(* IEC 61131-3 sources: volt/packages/volt-lsp-iec/test-corpus/awa-palletizer/Device/Plc Logic/Application/Library Manager/L_UMTP_Mathematics, 222 files *)

(* ---- L_UMTP_COMPLEX.dut ---- *)
TYPE L_UMTP_COMPLEX :
STRUCT
	LRRE : LREAL;
	LRIM : LREAL;
END_STRUCT
END_TYPE

(* ---- L_UMTP_INTERPOLATIONDATA.dut ---- *)
TYPE L_UMTP_INTERPOLATIONDATA :
STRUCT
	PARRX : POINTER TO LREAL;
	XISEQUIDISTANT : BOOL;
	UDISTRIDEX : UDINT;
	PARRY : POINTER TO LREAL;
	YISEQUIDISTANT : BOOL;
	UDISTRIDEY : UDINT;
	UICOUNT : UDINT;
	OPTIONS : UDINT;
END_STRUCT
END_TYPE

(* ---- L_UMTP_INTERPOLATIONTYPE.dut ---- *)
TYPE L_UMTP_INTERPOLATIONTYPE :
(
	UNDEFINED := 0,
	LINEAR := 1,
	CUBICSPLINENATURAL := 30,
	CUBICSPLINEHERMITE := 31,
	CUBICSPLINEHERMITEEXTERN := 32,
	NEWTON := 5
);
END_TYPE

(* ---- L_UMTP_MATRIX3X3.dut ---- *)
TYPE L_UMTP_MATRIX3X3 :
STRUCT
	M11 : LREAL;
	M12 : LREAL;
	M13 : LREAL;
	M21 : LREAL;
	M22 : LREAL;
	M23 : LREAL;
	M31 : LREAL;
	M32 : LREAL;
	M33 : LREAL;
END_STRUCT
END_TYPE

(* ---- L_UMTP_QUATERNION.dut ---- *)
TYPE L_UMTP_QUATERNION :
STRUCT
	LRRE : LREAL;
	LRIM1 : LREAL;
	LRIM2 : LREAL;
	LRIM3 : LREAL;
END_STRUCT
END_TYPE

(* ---- L_UMTP_REVERSEPOLISHNOTATIONTOKEN.dut ---- *)
TYPE L_UMTP_REVERSEPOLISHNOTATIONTOKEN :
(
	NONE := 0,
	PARENTHESIS := 1,
	FLOAT := 2,
	BOOLEAN := 3,
	NEGOTIATE := 4,
	PLUS := 10,
	MINUS := 11,
	MULTIPLIKATION := 12,
	DIVISION := 13,
	POW := 14,
	MODULO := 15,
	SINE := 20,
	COSINE := 21,
	TANGENS := 22,
	ASINE := 23,
	ACOSINE := 24,
	ATANGENS := 25,
	EXPONENTIAL := 40,
	LOGN := 41,
	LOG10 := 42,
	SQUAREROOT := 43,
	ABSOLUTE := 44,
	SIGNUM := 45,
	CEIL := 50,
	FLOOR := 51,
	TRUNCATE := 52,
	ROUND := 53,
	EQUAL := 100,
	NOTEQUAL := 101,
	GREATEREQUAL := 102,
	GREATERTHEN := 103,
	LESSEQUAL := 104,
	LESSTHEN := 105,
	LOGICAND := 110,
	LOGICXOR := 111,
	LOGICOR := 112,
	LOGICNOT := 113
);
END_TYPE

(* ---- L_UMTP_ROBOTACC.dut ---- *)
TYPE L_UMTP_ROBOTACC :
STRUCT
	ACC : L_UMTP_Vector3D;
	PITCH : L_UMTP_Vector3D;
END_STRUCT
END_TYPE

(* ---- L_UMTP_ROBOTFRAME.dut ---- *)
TYPE L_UMTP_ROBOTFRAME :
STRUCT
	POS : L_UMTP_RobotPos;
	VEL : L_UMTP_RobotVel;
	ACC : L_UMTP_RobotAcc;
END_STRUCT
END_TYPE

(* ---- L_UMTP_ROBOTPOS.dut ---- *)
TYPE L_UMTP_ROBOTPOS :
STRUCT
	POS : L_UMTP_Vector3D;
	ROT : L_UMTP_RotMat;
END_STRUCT
END_TYPE

(* ---- L_UMTP_ROBOTVEL.dut ---- *)
TYPE L_UMTP_ROBOTVEL :
STRUCT
	VEL : L_UMTP_Vector3D;
	TWIST : L_UMTP_Vector3D;
END_STRUCT
END_TYPE

(* ---- L_UMTP_ROTATIONCONVENTION.dut ---- *)
TYPE L_UMTP_ROTATIONCONVENTION :
(
	XYZ_ROTATED := 0,
	ZYX_ROTATED := 1,
	XZY_ROTATED := 2,
	YZX_ROTATED := 3,
	YXZ_ROTATED := 4,
	ZXY_ROTATED := 5,
	XYZ_FIXED := 100,
	ZYX_FIXED := 101,
	XZY_FIXED := 102,
	YZX_FIXED := 103,
	YXZ_FIXED := 104,
	ZXY_FIXED := 105
);
END_TYPE

(* ---- L_UMTP_ROTMAT.dut ---- *)
TYPE L_UMTP_ROTMAT :
STRUCT
	PARAM : L_UMTP_RotParam;
END_STRUCT
END_TYPE

(* ---- L_UMTP_ROTPARAM.dut ---- *)
TYPE L_UMTP_ROTPARAM :
STRUCT
	SINA : LREAL;
	COSA : LREAL;
	SINB : LREAL;
	COSB : LREAL;
	SINC : LREAL;
	COSC : LREAL;
	EROTCON : L_UMTP_RotationConvention;
	XGIMBALLOCK : BOOL;
END_STRUCT
END_TYPE

(* ---- L_UMTP_TRIGONOMETRICUNIT.dut ---- *)
TYPE L_UMTP_TRIGONOMETRICUNIT :
(
	RADIANT := 0,
	DEGREE := 1
);
END_TYPE

(* ---- L_UMTP_VALIDLREAL.dut ---- *)
TYPE L_UMTP_VALIDLREAL :
STRUCT
	XVALID : BOOL;
	LRVALUE : LREAL;
END_STRUCT
END_TYPE

(* ---- L_UMTP_VECTOR3D.dut ---- *)
TYPE L_UMTP_VECTOR3D :
STRUCT
	X : LREAL;
	Y : LREAL;
	Z : LREAL;
END_STRUCT
END_TYPE

(* ---- L_UMTP_CONSTANTS.gvl ---- *)
VAR_GLOBAL
	GC_CTRLPTMAXNR : INT := 200;
	GC_IMAXNUMOFGIVENPTS : INT := 199;
	GC_UDIMAXCUBSPLINEPTS : UDINT := 11;
	G_MAXPATHDIM : DINT := 8;
	GCDWSIZEOFLREAL : DWORD := USINT_TO_DWORD(SIZEOF(LREAL));
END_VAR

(* ---- L_UMTP_DEFINES.gvl ---- *)
VAR_GLOBAL
	G_XOPTIMIZEDFRAMECALC : BOOL := TRUE;
END_VAR

(* ---- L_UMTP_MATH.gvl ---- *)
VAR_GLOBAL
	RAD2DEG : LREAL := (180.0 / Math.PI);
	DEG2RAD : LREAL := (Math.PI / 180.0);
	GRAVITY_MM : LREAL := (9.81 * 1000.0);
	EPS_REAL : LREAL := 1E-06;
	GC_LREPSILON : LREAL := 1E-09;
	EPS_LREAL : LREAL := 1E-12;
	MM2M : LREAL := 0.001;
	M2MM : LREAL := 1000;
	GCGIMBALLOCKTOL : LREAL := 5E-05;
	GCLRINVPI : LREAL := (1 / MATH.PI);
	GCLR2PI : LREAL := (2 * MATH.PI);
	GCLRINV2PI : LREAL := (1 / (2 * MATH.PI));
	GCLRPIHALF : LREAL := (MATH.PI / 2);
	GCLRINVPIHALF : LREAL := (1 / (MATH.PI / 2));
	MAXDOUBLE : LREAL := 1.79769E+308;
	MINDOUBLE : LREAL := -1.79769E+308;
	GC_POSITIVE_LIMIT_16BIT_LREAL : LREAL := 65535.0;
	GC_POSITIVE_LIMIT_15BIT_LREAL : LREAL := 32767.0;
	GC_NEGATIVE_LIMIT_15BIT_LREAL : LREAL := -32768.0;
	GC_POSITIVE_LIMIT_32BIT : LREAL := 2147483647;
	GC_NEGATIVE_LIMIT_32BIT : LREAL := -2147483647;
	GC_POSITIVE_LIMIT_32BIT_LREAL : LREAL := 4294967296.0;
	GC_POSITIVE_LIMIT_31BIT_LREAL : LREAL := 2147483647.0;
	GC_NEGATIVE_LIMIT_31BIT_LREAL : LREAL := -2147483648.0;
	GC_POSITIVE_LIMIT_63BIT_LREAL : LREAL := 9.2233720368547758E+18;
	GC_NEGATIVE_LIMIT_63BIT_LREAL : LREAL := -9.2233720368547758E+18;
	GC_POSITIVE_LIMIT_63BIT : LINT := 9223372036854775807;
	GC_NEGATIVE_LIMIT_63BIT : LINT := -9223372036854775808;
	LRCOS_0 : LREAL := 1.0;
	LRCOS_15 : LREAL := 0.965925826289068;
	LRCOS_30 : LREAL := 0.866025403784439;
	LRCOS_45 : LREAL := 0.707106781186547;
	LRCOS_60 : LREAL := 0.5;
	LRCOS_75 : LREAL := 0.258819045102521;
	LRCOS_90 : LREAL := 0.0;
	LRCOS_105 : LREAL := -0.258819045102521;
	LRCOS_120 : LREAL := -0.5;
	LRCOS_135 : LREAL := -0.707106781186548;
	LRCOS_150 : LREAL := -0.866025403784439;
	LRCOS_165 : LREAL := -0.965925826289068;
	LRCOS_180 : LREAL := -1.0;
	LRCOS_195 : LREAL := -0.965925826289068;
	LRCOS_210 : LREAL := -0.866025403784439;
	LRCOS_225 : LREAL := -0.707106781186547;
	LRCOS_240 : LREAL := -0.5;
	LRCOS_255 : LREAL := -0.258819045102521;
	LRCOS_270 : LREAL := 0.0;
	LRCOS_285 : LREAL := 0.258819045102521;
	LRCOS_300 : LREAL := 0.5;
	LRCOS_315 : LREAL := 0.707106781186548;
	LRCOS_330 : LREAL := 0.866025403784439;
	LRCOS_345 : LREAL := 0.965925826289068;
	LRCOS_360 : LREAL := 1.0;
	LRSIN_0 : LREAL := 0.0;
	LRSIN_15 : LREAL := 0.258819045102521;
	LRSIN_30 : LREAL := 0.5;
	LRSIN_45 : LREAL := 0.707106781186548;
	LRSIN_60 : LREAL := 0.866025403784439;
	LRSIN_75 : LREAL := 0.965925826289068;
	LRSIN_90 : LREAL := 1.0;
	LRSIN_105 : LREAL := 0.965925826289068;
	LRSIN_120 : LREAL := 0.866025403784439;
	LRSIN_135 : LREAL := 0.707106781186547;
	LRSIN_150 : LREAL := 0.5;
	LRSIN_165 : LREAL := 0.258819045102521;
	LRSIN_180 : LREAL := 0.0;
	LRSIN_195 : LREAL := -0.258819045102521;
	LRSIN_210 : LREAL := -0.5;
	LRSIN_225 : LREAL := -0.707106781186548;
	LRSIN_240 : LREAL := -0.866025403784439;
	LRSIN_255 : LREAL := -0.965925826289068;
	LRSIN_270 : LREAL := -1.0;
	LRSIN_285 : LREAL := -0.965925826289068;
	LRSIN_300 : LREAL := -0.866025403784439;
	LRSIN_315 : LREAL := -0.707106781186547;
	LRSIN_330 : LREAL := -0.5;
	LRSIN_345 : LREAL := -0.258819045102521;
	LRSIN_360 : LREAL := 0.0;
	L_UMTP_VALUEIGNORE : LREAL := 1E+300;
	L_UMTP_VALUEINITIAL : LREAL := 1E+301;
	L_UMTP_VALUEINVALID : LREAL := 1E+302;
	L_UMTP_VALUEINF : LREAL := 1.7976931348623157E+308;
END_VAR

(* ---- L_UMTP_FUNC_1D21D.itf ---- *)
INTERFACE L_UMTP_FUNC_1D21D
END_INTERFACE

METHOD CALL_1D21D : LREAL
VAR_INPUT
	X : LREAL;
	CONTEXT : DINT;
END_VAR
END_METHOD

(* ---- L_UMTP_FUNC_ND21D.itf ---- *)
INTERFACE L_UMTP_FUNC_ND21D
END_INTERFACE

METHOD CALL_ND21D : LREAL
VAR_INPUT
	PLRX : POINTER TO LREAL;
	UDIDIM : UDINT;
	CONTEXT : DINT;
END_VAR
END_METHOD

(* ---- L_UMTP_FUNC_ND2MD.itf ---- *)
INTERFACE L_UMTP_FUNC_ND2MD
END_INTERFACE

METHOD CALL_ND2MD
VAR_INPUT
	PLRX : POINTER TO LREAL;
	UDIXDIM : UDINT;
	PLRY : POINTER TO LREAL;
	UDIYDIM : UDINT;
	CONTEXT : DINT;
END_VAR
END_METHOD

(* ---- L_UMTP_IFFTDATA.itf ---- *)
INTERFACE L_UMTP_IFFTDATA
END_INTERFACE

METHOD RECORDDATA : UDINT
VAR_INPUT
	PLCDATA : POINTER TO L_umtp_complex;
	UDISIZEOFDATA : UDINT;
END_VAR
END_METHOD

METHOD STARTRECORDING : BOOL
END_METHOD

METHOD STOPRECORDING : BOOL
END_METHOD

(* ---- L_UMTP_IINTERPOLATION.itf ---- *)
INTERFACE L_UMTP_IINTERPOLATION
END_INTERFACE

METHOD GETVALUE : BOOL
VAR_INPUT
	X : LREAL;
END_VAR
VAR_OUTPUT
	Y : LREAL;
END_VAR
END_METHOD

(* ---- L_UMTP_IMETRIC.itf ---- *)
INTERFACE L_UMTP_IMETRIC
END_INTERFACE

METHOD DISTANCE : LREAL
VAR_INPUT
	ITFOB1 : __SYSTEM.IQueryInterface;
	ITFOB2 : __SYSTEM.IQueryInterface;
END_VAR
END_METHOD

(* ---- L_UMTP_IODE.itf ---- *)
INTERFACE L_UMTP_IODE
END_INTERFACE

METHOD FIRSTDERIV
VAR_INPUT
	PLRY : POINTER TO LREAL;
	PLRDY : POINTER TO LREAL;
	UDIDIM : UDINT;
	LRT : LREAL;
END_VAR
END_METHOD

(* ---- L_UMTP_IPATH.itf ---- *)
INTERFACE L_UMTP_IPATH
END_INTERFACE

METHOD GETPATHVALUE : BOOL
VAR_INPUT
	PLRX : POINTER TO LREAL;
	PLRD1 : POINTER TO LREAL;
	PLRD2 : POINTER TO LREAL;
	UDIDIM : UDINT;
	LRU : LREAL;
END_VAR
END_METHOD

(* ---- L_UMTP_ISORTDATA.itf ---- *)
INTERFACE L_UMTP_ISORTDATA
END_INTERFACE

METHOD EXCHANGE : BOOL
VAR_INPUT
	IDX1 : DINT;
	IDX2 : DINT;
END_VAR
END_METHOD

METHOD GETVALUE : LREAL
VAR_INPUT
	IDX : DINT;
END_VAR
END_METHOD

(* ---- CALCCARTLENGTH.pou ---- *)
FUNCTION CALCCARTLENGTH : LREAL
VAR_INPUT
	PVEC : POINTER TO LREAL;
	NUMELEMENTS : __XWORD;
END_VAR
END_FUNCTION

(* ---- CAPITAL_CASE.pou ---- *)
FUNCTION CAPITAL_CASE : STRING(255)
VAR_INPUT
	STR : STRING(255);
END_VAR
END_FUNCTION

(* ---- DELETE_FROM_STR.pou ---- *)
FUNCTION DELETE_FROM_STR : STRING(255)
VAR_INPUT
	STR1 : STRING(255);
	STR2 : STRING(255);
END_VAR
END_FUNCTION

(* ---- GETBOOLEANPROPERTY.pou ---- *)
FUNCTION GETBOOLEANPROPERTY : BOOL
VAR_INPUT
	STKEY : WSTRING;
END_VAR
END_FUNCTION

(* ---- GETCOMPANY.pou ---- *)
FUNCTION GETCOMPANY : WSTRING
END_FUNCTION

(* ---- GETNUMBERPROPERTY.pou ---- *)
FUNCTION GETNUMBERPROPERTY : DINT
VAR_INPUT
	STKEY : WSTRING;
END_VAR
END_FUNCTION

(* ---- GETTEXTPROPERTY.pou ---- *)
FUNCTION GETTEXTPROPERTY : WSTRING
VAR_INPUT
	STKEY : WSTRING;
END_VAR
END_FUNCTION

(* ---- GETTEXTPROPERTY2.pou ---- *)
FUNCTION GETTEXTPROPERTY2 : POINTER TO WSTRING
VAR_INPUT
	STKEY : WSTRING;
END_VAR
END_FUNCTION

(* ---- GETTITLE.pou ---- *)
FUNCTION GETTITLE : WSTRING
END_FUNCTION

(* ---- GETVERSION.pou ---- *)
FUNCTION GETVERSION : VERSION
END_FUNCTION

(* ---- GETVERSIONPROPERTY.pou ---- *)
FUNCTION GETVERSIONPROPERTY : VERSION
VAR_INPUT
	STKEY : WSTRING;
END_VAR
END_FUNCTION

(* ---- L_UMTP_2DINTERPOLATIONLINEAR.pou ---- *)
FUNCTION L_UMTP_2DINTERPOLATIONLINEAR : BOOL
VAR_INPUT
	ALRX : POINTER TO LREAL;
	ALRY : POINTER TO LREAL;
	ALRZ : POINTER TO LREAL;
	LRX : LREAL;
	LRY : LREAL;
END_VAR
VAR_OUTPUT
	XERROR : BOOL;
	EERRORID : L_IE1P_Error;
	LRZ : LREAL;
END_VAR
END_FUNCTION

(* ---- L_UMTP_ABC2ROT.pou ---- *)
FUNCTION L_UMTP_ABC2ROT
VAR_INPUT
	ROTMAT : REFERENCE TO L_UMTP_RotMat;
END_VAR
END_FUNCTION

(* ---- L_UMTP_ANTISYMTIMESMATRIX3D.pou ---- *)
FUNCTION L_UMTP_ANTISYMTIMESMATRIX3D
VAR_INPUT
	M : REFERENCE TO L_UMTP_Matrix3x3;
	TWIST : REFERENCE TO L_UMTP_Vector3D;
	RESULT : REFERENCE TO L_UMTP_Matrix3x3;
END_VAR
END_FUNCTION

(* ---- L_UMTP_APPENDPITCH.pou ---- *)
FUNCTION L_UMTP_APPENDPITCH : BOOL
VAR_INPUT
	DPHIA : LREAL;
	DPHIB : LREAL;
	DPHIC : LREAL;
	DDPHIA : LREAL;
	DDPHIB : LREAL;
	DDPHIC : LREAL;
	FRAME : REFERENCE TO L_UMTP_RobotFrame;
END_VAR
END_FUNCTION

(* ---- L_UMTP_APPENDTWIST.pou ---- *)
FUNCTION L_UMTP_APPENDTWIST : BOOL
VAR_INPUT
	DPHIA : LREAL;
	DPHIB : LREAL;
	DPHIC : LREAL;
	FRAME : REFERENCE TO L_UMTP_RobotFrame;
END_VAR
END_FUNCTION

(* ---- L_UMTP_APPROXSIGN.pou ---- *)
FUNCTION L_UMTP_APPROXSIGN : LREAL
VAR_INPUT
	LRX : LREAL;
	LRFAC : LREAL;
END_VAR
END_FUNCTION

(* ---- L_UMTP_ATAN2.pou ---- *)
FUNCTION L_UMTP_ATAN2 : LREAL
VAR_INPUT
	LRSINUS : LREAL;
	LRCOSINUS : LREAL;
END_VAR
END_FUNCTION

(* ---- L_UMTP_BENDING.pou ---- *)
FUNCTION L_UMTP_BENDING : LREAL
VAR_INPUT
	ALRD1 : REFERENCE TO ARRAY [1..3] OF LREAL;
	ALRD2 : REFERENCE TO ARRAY [1..3] OF LREAL;
END_VAR
END_FUNCTION

(* ---- L_UMTP_BILINEARINTERPOLATION.pou ---- *)
FUNCTION L_UMTP_BILINEARINTERPOLATION : BOOL
VAR_INPUT
	LRX0 : LREAL;
	LRX1 : LREAL;
	LRY0 : LREAL;
	LRY1 : LREAL;
	LRZ00 : LREAL;
	LRZ01 : LREAL;
	LRZ10 : LREAL;
	LRZ11 : LREAL;
	LRX : LREAL;
	LRY : LREAL;
END_VAR
VAR_OUTPUT
	LRZ : LREAL;
END_VAR
END_FUNCTION

(* ---- L_UMTP_BISECTION.pou ---- *)
FUNCTION L_UMTP_BISECTION : BOOL
VAR_INPUT
	IFUNC : L_UMTP_Func_1D21D;
	CONTEXT : DINT;
	A : LREAL;
	B : LREAL;
	F_REQUESTED : LREAL;
	TOL : LREAL;
	X : REFERENCE TO LREAL;
END_VAR
END_FUNCTION

(* ---- L_UMTP_BRENTALGORITHM.pou ---- *)
FUNCTION L_UMTP_BRENTALGORITHM : BOOL
VAR_INPUT
	IFUNC : L_UMTP_Func_1D21D;
	CONTEXT : DINT;
	A : LREAL;
	B : LREAL;
	TOL : LREAL;
	X : REFERENCE TO LREAL;
END_VAR
END_FUNCTION

(* ---- L_UMTP_BUBBLESORTINT.pou ---- *)
FUNCTION L_UMTP_BUBBLESORTINT
VAR_INPUT
	PIX : POINTER TO INT;
	UDISIZE : UDINT;
	XINVERT : BOOL;
END_VAR
END_FUNCTION

(* ---- L_UMTP_BUBBLESORTITFSORTDATA.pou ---- *)
FUNCTION L_UMTP_BUBBLESORTITFSORTDATA : BOOL
VAR_INPUT
	ITFDATA : L_UMTP_ISortData;
	XINVERT : BOOL;
END_VAR
END_FUNCTION

(* ---- L_UMTP_BUBBLESORTLREAL.pou ---- *)
FUNCTION L_UMTP_BUBBLESORTLREAL
VAR_INPUT
	PLRX : POINTER TO LREAL;
	UDISIZE : UDINT;
	XINVERT : BOOL;
END_VAR
END_FUNCTION

(* ---- L_UMTP_CHECKGIMBALLOCK.pou ---- *)
FUNCTION L_UMTP_CHECKGIMBALLOCK : BOOL
VAR_INPUT
	PARAM : REFERENCE TO L_UMTP_RotParam;
END_VAR
END_FUNCTION

(* ---- L_UMTP_CHECKMONOTONIC.pou ---- *)
FUNCTION L_UMTP_CHECKMONOTONIC : BYTE
VAR_INPUT
	PLRVALUES : POINTER TO LREAL;
	NDATA : UDINT;
	NSTRIDE : UDINT;
END_VAR
END_FUNCTION

(* ---- L_UMTP_CHECKSTEPSIZE.pou ---- *)
FUNCTION L_UMTP_CHECKSTEPSIZE : BOOL
VAR_INPUT
	PLRY0 : POINTER TO LREAL;
	PLRY1 : POINTER TO LREAL;
	UDIDIM : UDINT;
	LRTOL : LREAL;
	LRH : LREAL;
END_VAR
VAR_OUTPUT
	LRHTOL : LREAL;
END_VAR
END_FUNCTION

(* ---- L_UMTP_CLEAR.pou ---- *)
FUNCTION L_UMTP_CLEAR : BOOL
VAR_INPUT
	ALRARR : POINTER TO LREAL;
END_VAR
END_FUNCTION

(* ---- L_UMTP_COMEQ.pou ---- *)
FUNCTION L_UMTP_COMEQ : BOOL
VAR_INPUT
	COMVALUE : L_UMTP_Complex;
	COMTARGET : L_UMTP_Complex;
END_VAR
END_FUNCTION

(* ---- L_UMTP_COMPLEX2MAGNITUDE.pou ---- *)
FUNCTION L_UMTP_COMPLEX2MAGNITUDE : LREAL
VAR_INPUT
	SCCOIN : L_UMTP_Complex;
END_VAR
END_FUNCTION

(* ---- L_UMTP_COMPLEXCART2POLAR.pou ---- *)
FUNCTION L_UMTP_COMPLEXCART2POLAR
VAR_INPUT
	SCCOIN : L_UMTP_Complex;
	ETRIGUNIT : L_UMTP_TrigonometricUnit;
END_VAR
VAR_OUTPUT
	LRMAGNITUDE : LREAL;
	LRANGLE : LREAL;
END_VAR
END_FUNCTION

(* ---- L_UMTP_COMPLEXDIV.pou ---- *)
FUNCTION L_UMTP_COMPLEXDIV : L_UMTP_Complex
VAR_INPUT
	SCCOIN1 : L_UMTP_complex;
	SCCOIN2 : L_UMTP_complex;
END_VAR
END_FUNCTION

(* ---- L_UMTP_COMPLEXMUL.pou ---- *)
FUNCTION L_UMTP_COMPLEXMUL : L_UMTP_Complex
VAR_INPUT
	COIN1 : L_UMTP_complex;
	COIN2 : L_UMTP_complex;
END_VAR
END_FUNCTION

(* ---- L_UMTP_COMPLEXPOLAR2CART.pou ---- *)
FUNCTION L_UMTP_COMPLEXPOLAR2CART : L_UMTP_Complex
VAR_INPUT
	LRMAGNITUDE : LREAL;
	LRANGLE : LREAL;
	ETRIGUNIT : L_UMTP_TrigonometricUnit;
END_VAR
END_FUNCTION

(* ---- L_UMTP_CONFIGURATIONABC.pou ---- *)
FUNCTION L_UMTP_CONFIGURATIONABC : INT
VAR_INPUT
	ROTMAT : REFERENCE TO L_UMTP_RotMat;
END_VAR
END_FUNCTION

(* ---- L_UMTP_CROSS.pou ---- *)
FUNCTION L_UMTP_CROSS : BOOL
VAR_INPUT
	A : REFERENCE TO ARRAY [1..3] OF LREAL;
	B : REFERENCE TO ARRAY [1..3] OF LREAL;
	RESULT : REFERENCE TO ARRAY [1..3] OF LREAL;
END_VAR
END_FUNCTION

(* ---- L_UMTP_CROSSPROD.pou ---- *)
FUNCTION L_UMTP_CROSSPROD : BOOL
VAR_IN_OUT
	ALRA : ARRAY [1..3] OF LREAL;
	ALRB : ARRAY [1..3] OF LREAL;
	ALRRESULT : ARRAY [1..3] OF LREAL;
END_VAR
END_FUNCTION

(* ---- L_UMTP_DABC2DROT.pou ---- *)
FUNCTION L_UMTP_DABC2DROT
VAR_INPUT
	PARAM : REFERENCE TO L_UMTP_RotParam;
	DPHIA : LREAL;
	DPHIB : LREAL;
	DPHIC : LREAL;
	DROT : REFERENCE TO L_UMTP_Matrix3x3;
END_VAR
END_FUNCTION

(* ---- L_UMTP_DDABC2DDROT.pou ---- *)
FUNCTION L_UMTP_DDABC2DDROT
VAR_INPUT
	PARAM : L_UMTP_RotParam;
	DPHIA : LREAL;
	DPHIB : LREAL;
	DPHIC : LREAL;
	DDPHIA : LREAL;
	DDPHIB : LREAL;
	DDPHIC : LREAL;
	DDROT : REFERENCE TO L_UMTP_Matrix3x3;
END_VAR
END_FUNCTION

(* ---- L_UMTP_DDROT2DDABC.pou ---- *)
FUNCTION L_UMTP_DDROT2DDABC
VAR_INPUT
	PARAM : REFERENCE TO L_UMTP_RotParam;
	DDROT : REFERENCE TO L_UMTP_Matrix3x3;
	DPHIA : LREAL;
	DPHIB : LREAL;
	DPHIC : LREAL;
END_VAR
VAR_OUTPUT
	DDPHIA : LREAL;
	DDPHIB : LREAL;
	DDPHIC : LREAL;
END_VAR
END_FUNCTION

(* ---- L_UMTP_DDROT2FRAME.pou ---- *)
FUNCTION L_UMTP_DDROT2FRAME : BOOL
VAR_INPUT
	FRAME : REFERENCE TO L_UMTP_RobotFrame;
	DDROT : REFERENCE TO L_UMTP_Matrix3x3;
END_VAR
END_FUNCTION

(* ---- L_UMTP_DETERMINAT3D.pou ---- *)
FUNCTION L_UMTP_DETERMINAT3D : LREAL
VAR_IN_OUT
	M : L_UMTP_Matrix3x3;
END_VAR
END_FUNCTION

(* ---- L_UMTP_DISTANCE.pou ---- *)
FUNCTION L_UMTP_DISTANCE : LREAL
VAR_INPUT
	PLRX : POINTER TO LREAL;
	PLRY : POINTER TO LREAL;
	UDIDIM : UDINT;
END_VAR
END_FUNCTION

(* ---- L_UMTP_DIV.pou ---- *)
FUNCTION L_UMTP_DIV : LREAL
VAR_INPUT
	A : LREAL;
	B : LREAL;
END_VAR
END_FUNCTION

(* ---- L_UMTP_DORMANDPRINCE45STEP.pou ---- *)
FUNCTION L_UMTP_DORMANDPRINCE45STEP
VAR_INPUT
	IODE : L_UMTP_IODE;
	PLRY0 : POINTER TO LREAL;
	UDIDIM : UDINT;
	LRT : LREAL;
	LRH : LREAL;
	LRTOL : LREAL;
END_VAR
VAR_OUTPUT
	LRTNEW : LREAL;
	XACCEPTED : BOOL;
	UDIREPEATS : UDINT;
END_VAR
END_FUNCTION

(* ---- L_UMTP_DROT2DABC.pou ---- *)
FUNCTION L_UMTP_DROT2DABC
VAR_INPUT
	PARAM : REFERENCE TO L_UMTP_RotParam;
	DROT : REFERENCE TO L_UMTP_Matrix3x3;
END_VAR
VAR_OUTPUT
	DPHIA : LREAL;
	DPHIB : LREAL;
	DPHIC : LREAL;
END_VAR
END_FUNCTION

(* ---- L_UMTP_DROT2FRAME.pou ---- *)
FUNCTION L_UMTP_DROT2FRAME : BOOL
VAR_INPUT
	FRAME : REFERENCE TO L_UMTP_RobotFrame;
	DROT : REFERENCE TO L_UMTP_Matrix3x3;
END_VAR
END_FUNCTION

(* ---- L_UMTP_ENSURE180.pou ---- *)
FUNCTION L_UMTP_ENSURE180 : LREAL
VAR_INPUT
	LRVALUE : LREAL;
END_VAR
VAR_OUTPUT
	IINTERVALCOUNT : LINT;
END_VAR
END_FUNCTION

(* ---- L_UMTP_ENSUREINTERVAL.pou ---- *)
FUNCTION L_UMTP_ENSUREINTERVAL : LREAL
VAR_INPUT
	LRVALUE : LREAL;
	LRLOWER : LREAL;
	LRUPPER : LREAL;
END_VAR
VAR_OUTPUT
	IINTERVALCOUNT : LINT;
END_VAR
END_FUNCTION

(* ---- L_UMTP_ENSUREMAXDIFF360.pou ---- *)
FUNCTION L_UMTP_ENSUREMAXDIFF360 : LREAL
VAR_INPUT
	LRVALUE : LREAL;
	LRREFERENCE : LREAL;
	LRDIFF : LREAL;
END_VAR
VAR_OUTPUT
	IINTERVALCOUNT : LINT;
	XERROR : BOOL;
END_VAR
END_FUNCTION

(* ---- L_UMTP_ENSUREPI.pou ---- *)
FUNCTION L_UMTP_ENSUREPI : LREAL
VAR_INPUT
	LRVALUE : LREAL;
END_VAR
VAR_OUTPUT
	IINTERVALCOUNT : LINT;
END_VAR
END_FUNCTION

(* ---- L_UMTP_EULERSTEP.pou ---- *)
FUNCTION L_UMTP_EULERSTEP
VAR_INPUT
	IODE : L_UMTP_IODE;
	PLRY0 : POINTER TO LREAL;
	UDIDIM : UDINT;
	LRT : LREAL;
	LRH : LREAL;
END_VAR
VAR_OUTPUT
	LRTNEW : LREAL;
END_VAR
END_FUNCTION

(* ---- L_UMTP_EXPTAYLOR.pou ---- *)
FUNCTION L_UMTP_EXPTAYLOR : LREAL
VAR_INPUT
	LRX : LREAL;
END_VAR
END_FUNCTION

(* ---- L_UMTP_EXTRAPOLATEFRAME.pou ---- *)
FUNCTION L_UMTP_EXTRAPOLATEFRAME : BOOL
VAR_INPUT
	LRTIME : LREAL;
END_VAR
VAR_IN_OUT
	SCFRAME : L_UMTP_RobotFrame;
END_VAR
END_FUNCTION

(* ---- L_UMTP_FADFRAME.pou ---- *)
FUNCTION L_UMTP_FADFRAME : BOOL
VAR_INPUT
	LRFADFACTOR : LREAL;
END_VAR
VAR_IN_OUT
	SCFRAME : L_UMTP_RobotFrame;
	SCROTVECTOR : L_UMTP_Vector3D;
	SCFRAMEFADED : L_UMTP_RobotFrame;
	SCROTVECTORFADED : L_UMTP_Vector3D;
END_VAR
END_FUNCTION

(* ---- L_UMTP_FINDINTERVAL.pou ---- *)
FUNCTION L_UMTP_FINDINTERVAL : BOOL
VAR_INPUT
	LRVALUE : LREAL;
	PLRVALUES : POINTER TO LREAL;
	NDATA : UDINT;
	NSTRIDE : UDINT;
	XTRYFIRST : BOOL;
END_VAR
VAR_OUTPUT
	XERROR : BOOL;
	EERRORID : L_IE1P_Error;
END_VAR
VAR_IN_OUT
	UDIINTERVAL : UDINT;
END_VAR
END_FUNCTION

(* ---- L_UMTP_FRAME2DDROT.pou ---- *)
FUNCTION L_UMTP_FRAME2DDROT : BOOL
VAR_INPUT
	FRAME : REFERENCE TO L_UMTP_RobotFrame;
	DDROT : REFERENCE TO L_UMTP_Matrix3x3;
END_VAR
END_FUNCTION

(* ---- L_UMTP_FRAME2DROT.pou ---- *)
FUNCTION L_UMTP_FRAME2DROT : BOOL
VAR_INPUT
	FRAME : REFERENCE TO L_UMTP_RobotFrame;
	DROT : REFERENCE TO L_UMTP_Matrix3x3;
END_VAR
END_FUNCTION

(* ---- L_UMTP_FRAMETIMESFRAME.pou ---- *)
FUNCTION L_UMTP_FRAMETIMESFRAME
VAR_INPUT
	FRAMEA : REFERENCE TO L_UMTP_RobotFrame;
	FRAMEB : REFERENCE TO L_UMTP_RobotFrame;
	RESULT : REFERENCE TO L_UMTP_RobotFrame;
END_VAR
END_FUNCTION

(* ---- L_UMTP_FRAMETIMESFRAMEACC.pou ---- *)
FUNCTION L_UMTP_FRAMETIMESFRAMEACC : BOOL
VAR_INPUT
	FRAMEA : REFERENCE TO L_UMTP_RobotFrame;
	FRAMEB : REFERENCE TO L_UMTP_RobotFrame;
	RESULT : REFERENCE TO L_UMTP_RobotFrame;
END_VAR
END_FUNCTION

(* ---- L_UMTP_FRAMETIMESFRAMEPOS.pou ---- *)
FUNCTION L_UMTP_FRAMETIMESFRAMEPOS
VAR_INPUT
	FRAMEA : REFERENCE TO L_UMTP_RobotFrame;
	FRAMEB : REFERENCE TO L_UMTP_RobotFrame;
	RESULT : REFERENCE TO L_UMTP_RobotFrame;
END_VAR
END_FUNCTION

(* ---- L_UMTP_FRAMETIMESFRAMEVEL.pou ---- *)
FUNCTION L_UMTP_FRAMETIMESFRAMEVEL : BOOL
VAR_INPUT
	FRAMEA : REFERENCE TO L_UMTP_RobotFrame;
	FRAMEB : REFERENCE TO L_UMTP_RobotFrame;
	RESULT : REFERENCE TO L_UMTP_RobotFrame;
END_VAR
END_FUNCTION

(* ---- L_UMTP_FRAMETIMESROBOTPOS.pou ---- *)
FUNCTION L_UMTP_FRAMETIMESROBOTPOS
VAR_INPUT
	FRAME : REFERENCE TO L_UMTP_RobotFrame;
	ROBOTPOS : REFERENCE TO L_UMTP_RobotPos;
	RESULT : REFERENCE TO L_UMTP_RobotFrame;
END_VAR
END_FUNCTION

(* ---- L_UMTP_FRAMETIMESROBOTPOSACC.pou ---- *)
FUNCTION L_UMTP_FRAMETIMESROBOTPOSACC
VAR_INPUT
	FRAME : REFERENCE TO L_UMTP_RobotFrame;
	ROBOTPOS : REFERENCE TO L_UMTP_RobotPos;
	RESULT : REFERENCE TO L_UMTP_RobotFrame;
END_VAR
END_FUNCTION

(* ---- L_UMTP_FRAMETIMESROBOTPOSPOS.pou ---- *)
FUNCTION L_UMTP_FRAMETIMESROBOTPOSPOS
VAR_INPUT
	FRAME : REFERENCE TO L_UMTP_RobotFrame;
	ROBOTPOS : REFERENCE TO L_UMTP_RobotPos;
	RESULT : REFERENCE TO L_UMTP_RobotFrame;
END_VAR
END_FUNCTION

(* ---- L_UMTP_FRAMETIMESROBOTPOSVEL.pou ---- *)
FUNCTION L_UMTP_FRAMETIMESROBOTPOSVEL
VAR_INPUT
	FRAME : REFERENCE TO L_UMTP_RobotFrame;
	ROBOTPOS : REFERENCE TO L_UMTP_RobotPos;
	RESULT : REFERENCE TO L_UMTP_RobotFrame;
END_VAR
END_FUNCTION

(* ---- L_UMTP_GENERATEROT.pou ---- *)
FUNCTION L_UMTP_GENERATEROT
VAR_INPUT
	SCTWIST : L_UMTP_Vector3D;
	LRTIME : LREAL;
END_VAR
VAR_IN_OUT
	SCROTRESULT : L_UMTP_RotMat;
END_VAR
END_FUNCTION

(* ---- L_UMTP_HLPINTERPOLATIONBILINEAREBETWEENLIMITS.pou ---- *)
FUNCTION L_UMTP_HLPINTERPOLATIONBILINEAREBETWEENLIMITS : LREAL
VAR_INPUT
	LRXSCALED : LREAL;
	LRYSCALED : LREAL;
END_VAR
VAR_IN_OUT
	ALRPAR2D : ARRAY [1..2, 1..2] OF LREAL;
END_VAR
END_FUNCTION

(* ---- L_UMTP_HLPINTERPOLATIONLINEARBETWEENLIMITS.pou ---- *)
FUNCTION L_UMTP_HLPINTERPOLATIONLINEARBETWEENLIMITS : LREAL
VAR_INPUT
	LRXSCALED : LREAL;
END_VAR
VAR_IN_OUT
	ALRPAR : ARRAY [1..2] OF LREAL;
END_VAR
END_FUNCTION

(* ---- L_UMTP_HOMMATRIXTOROBOTPOS.pou ---- *)
FUNCTION L_UMTP_HOMMATRIXTOROBOTPOS
VAR_INPUT
	HOMMATRIX : REFERENCE TO ARRAY [1..4, 1..4] OF LREAL;
	ROBOTPOS : REFERENCE TO L_UMTP_RobotPos;
	LRSCALEMATRIX2POS : LREAL;
END_VAR
END_FUNCTION

(* ---- L_UMTP_INVERT.pou ---- *)
FUNCTION L_UMTP_INVERT : BOOL
VAR_INPUT
	PLRM : POINTER TO LREAL;
	PLRMINV : POINTER TO LREAL;
	UDIROWS : UDINT;
	UDICOLS : UDINT;
END_VAR
END_FUNCTION

(* ---- L_UMTP_INVERT2X2.pou ---- *)
FUNCTION L_UMTP_INVERT2X2 : BOOL
VAR_IN_OUT
	ALRM : ARRAY [1..2, 1..2] OF LREAL;
	ALRMINV : ARRAY [1..2, 1..2] OF LREAL;
END_VAR
END_FUNCTION

(* ---- L_UMTP_INVERT3X3.pou ---- *)
FUNCTION L_UMTP_INVERT3X3 : BOOL
VAR_IN_OUT
	ALRM : ARRAY [1..3, 1..3] OF LREAL;
	ALRMINV : ARRAY [1..3, 1..3] OF LREAL;
END_VAR
END_FUNCTION

(* ---- L_UMTP_INVERTROBOTACC.pou ---- *)
FUNCTION L_UMTP_INVERTROBOTACC : BOOL
VAR_INPUT
	FRAME : REFERENCE TO L_UMTP_RobotFrame;
	FRAMEINV : REFERENCE TO L_UMTP_RobotFrame;
END_VAR
END_FUNCTION

(* ---- L_UMTP_INVERTROBOTFRAME.pou ---- *)
FUNCTION L_UMTP_INVERTROBOTFRAME : BOOL
VAR_INPUT
	FRAME : REFERENCE TO L_UMTP_RobotFrame;
	FRAMEINV : REFERENCE TO L_UMTP_RobotFrame;
END_VAR
END_FUNCTION

(* ---- L_UMTP_INVERTROBOTPOS.pou ---- *)
FUNCTION L_UMTP_INVERTROBOTPOS
VAR_INPUT
	ROBOTPOS : REFERENCE TO L_UMTP_RobotPos;
	ROBOTPOSINV : REFERENCE TO L_UMTP_RobotPos;
END_VAR
END_FUNCTION

(* ---- L_UMTP_INVERTROBOTVEL.pou ---- *)
FUNCTION L_UMTP_INVERTROBOTVEL : BOOL
VAR_INPUT
	FRAME : REFERENCE TO L_UMTP_RobotFrame;
	FRAMEINV : REFERENCE TO L_UMTP_RobotFrame;
END_VAR
END_FUNCTION

(* ---- L_UMTP_ISANTISYM.pou ---- *)
FUNCTION L_UMTP_ISANTISYM : BOOL
VAR_INPUT
	MAT : REFERENCE TO L_UMTP_Matrix3x3;
END_VAR
END_FUNCTION

(* ---- L_UMTP_ISIDENTITY.pou ---- *)
FUNCTION L_UMTP_ISIDENTITY : BOOL
VAR_INPUT
	M : REFERENCE TO L_UMTP_Matrix3x3;
END_VAR
END_FUNCTION

(* ---- L_UMTP_ISIDENTITYFRAME.pou ---- *)
FUNCTION L_UMTP_ISIDENTITYFRAME : BOOL
VAR_INPUT
	FRAME : REFERENCE TO L_UMTP_RobotFrame;
END_VAR
END_FUNCTION

(* ---- L_UMTP_ISNAN.pou ---- *)
FUNCTION L_UMTP_ISNAN : BOOL
VAR_INPUT
	LRVALUE : LREAL;
END_VAR
END_FUNCTION

(* ---- L_UMTP_ISSTATIONARYFRAME.pou ---- *)
FUNCTION L_UMTP_ISSTATIONARYFRAME : BOOL
VAR_INPUT
	FRAME : REFERENCE TO L_UMTP_RobotFrame;
END_VAR
END_FUNCTION

(* ---- L_UMTP_LINEARINTERPOLATION.pou ---- *)
FUNCTION L_UMTP_LINEARINTERPOLATION : BOOL
VAR_INPUT
	LRX0 : LREAL;
	LRX1 : LREAL;
	LRY0 : LREAL;
	LRY1 : LREAL;
	LRX : LREAL;
END_VAR
VAR_OUTPUT
	LRY : LREAL;
END_VAR
END_FUNCTION

(* ---- L_UMTP_LNTAYLOR.pou ---- *)
FUNCTION L_UMTP_LNTAYLOR : LREAL
VAR_INPUT
	LRY : LREAL;
END_VAR
END_FUNCTION

(* ---- L_UMTP_LREAL_TO_DINT.pou ---- *)
FUNCTION L_UMTP_LREAL_TO_DINT : DINT
VAR_INPUT
	LRVALUE : LREAL;
END_VAR
END_FUNCTION

(* ---- L_UMTP_LREAL_TO_DINT_TO_DWORD.pou ---- *)
FUNCTION L_UMTP_LREAL_TO_DINT_TO_DWORD : DWORD
VAR_INPUT
	LRVALUE : LREAL;
END_VAR
END_FUNCTION

(* ---- L_UMTP_LREAL_TO_DWORD.pou ---- *)
FUNCTION L_UMTP_LREAL_TO_DWORD : DWORD
VAR_INPUT
	LRVALUE : LREAL;
END_VAR
END_FUNCTION

(* ---- L_UMTP_LREAL_TO_INT.pou ---- *)
FUNCTION L_UMTP_LREAL_TO_INT : INT
VAR_INPUT
	LRVALUE : LREAL;
END_VAR
END_FUNCTION

(* ---- L_UMTP_LREAL_TO_INT_TO_WORD.pou ---- *)
FUNCTION L_UMTP_LREAL_TO_INT_TO_WORD : WORD
VAR_INPUT
	LRVALUE : LREAL;
END_VAR
END_FUNCTION

(* ---- L_UMTP_LREAL_TO_WORD.pou ---- *)
FUNCTION L_UMTP_LREAL_TO_WORD : WORD
VAR_INPUT
	LRVALUE : LREAL;
END_VAR
END_FUNCTION

(* ---- L_UMTP_LREQ.pou ---- *)
FUNCTION L_UMTP_LREQ : BOOL
VAR_INPUT
	LRVALUE : LREAL;
	LRTARGET : LREAL;
END_VAR
END_FUNCTION

(* ---- L_UMTP_LREQROT.pou ---- *)
FUNCTION L_UMTP_LREQROT : BOOL
VAR_INPUT
	LRA : LREAL;
	LRB : LREAL;
	LRC : LREAL;
	EROTCON : L_UMTP_RotationConvention;
	LRATARGET : LREAL;
	LRBTARGET : LREAL;
	LRCTARGET : LREAL;
	EROTCONTARGET : L_UMTP_RotationConvention;
END_VAR
END_FUNCTION

(* ---- L_UMTP_LRGE.pou ---- *)
FUNCTION L_UMTP_LRGE : BOOL
VAR_INPUT
	LRVALUE : LREAL;
	LRTARGET : LREAL;
END_VAR
END_FUNCTION

(* ---- L_UMTP_LRGT.pou ---- *)
FUNCTION L_UMTP_LRGT : BOOL
VAR_INPUT
	LRVALUE : LREAL;
	LRTARGET : LREAL;
END_VAR
END_FUNCTION

(* ---- L_UMTP_LRLE.pou ---- *)
FUNCTION L_UMTP_LRLE : BOOL
VAR_INPUT
	LRVALUE : LREAL;
	LRTARGET : LREAL;
END_VAR
END_FUNCTION

(* ---- L_UMTP_LRLT.pou ---- *)
FUNCTION L_UMTP_LRLT : BOOL
VAR_INPUT
	LRVALUE : LREAL;
	LRTARGET : LREAL;
END_VAR
END_FUNCTION

(* ---- L_UMTP_LRNE.pou ---- *)
FUNCTION L_UMTP_LRNE : BOOL
VAR_INPUT
	LRVALUE : LREAL;
	LRTARGET : LREAL;
END_VAR
END_FUNCTION

(* ---- L_UMTP_MATRIXADDMATRIX3D.pou ---- *)
FUNCTION L_UMTP_MATRIXADDMATRIX3D
VAR_INPUT
	A : REFERENCE TO L_UMTP_Matrix3x3;
	B : REFERENCE TO L_UMTP_Matrix3x3;
	RESULT : REFERENCE TO L_UMTP_Matrix3x3;
END_VAR
END_FUNCTION

(* ---- L_UMTP_MATRIXGET.pou ---- *)
FUNCTION L_UMTP_MATRIXGET : LREAL
VAR_INPUT
	I : UDINT;
	J : UDINT;
	STRIDE : UDINT;
	PMATRIX : POINTER TO LREAL;
END_VAR
END_FUNCTION

(* ---- L_UMTP_MATRIXINDEX.pou ---- *)
FUNCTION L_UMTP_MATRIXINDEX : UDINT
VAR_INPUT
	I : UDINT;
	J : UDINT;
	STRIDE : UDINT;
END_VAR
END_FUNCTION

(* ---- L_UMTP_MATRIXLN.pou ---- *)
FUNCTION L_UMTP_MATRIXLN : BOOL
VAR_IN_OUT
	SCROTMATRIX : L_UMTP_RotMat;
	SCROTVECTOR : L_UMTP_Vector3D;
END_VAR
END_FUNCTION

(* ---- L_UMTP_MATRIXSET.pou ---- *)
FUNCTION L_UMTP_MATRIXSET
VAR_INPUT
	I : UDINT;
	J : UDINT;
	STRIDE : UDINT;
	PMATRIX : POINTER TO LREAL;
	LRVALUE : LREAL;
END_VAR
END_FUNCTION

(* ---- L_UMTP_MATRIXTIMESANTISYM3D.pou ---- *)
FUNCTION L_UMTP_MATRIXTIMESANTISYM3D
VAR_INPUT
	M : REFERENCE TO L_UMTP_Matrix3x3;
	ASYM : REFERENCE TO L_UMTP_Vector3D;
	RESULT : REFERENCE TO L_UMTP_Matrix3x3;
END_VAR
END_FUNCTION

(* ---- L_UMTP_MATRIXTIMESMATRIX.pou ---- *)
FUNCTION L_UMTP_MATRIXTIMESMATRIX
VAR_INPUT
	PA : POINTER TO LREAL;
	PB : POINTER TO LREAL;
	PRESULT : POINTER TO LREAL;
	ZEILEN_A : __XWORD;
	SPALTEN_A : __XWORD;
	SPALTEN_B : __XWORD;
END_VAR
END_FUNCTION

(* ---- L_UMTP_MATRIXTIMESMATRIX3D.pou ---- *)
FUNCTION L_UMTP_MATRIXTIMESMATRIX3D
VAR_INPUT
	A : REFERENCE TO L_UMTP_Matrix3x3;
	B : REFERENCE TO L_UMTP_Matrix3x3;
	RESULT : REFERENCE TO L_UMTP_Matrix3x3;
END_VAR
END_FUNCTION

(* ---- L_UMTP_MATRIXTIMESMATRIXTRANSPOSE3D.pou ---- *)
FUNCTION L_UMTP_MATRIXTIMESMATRIXTRANSPOSE3D
VAR_INPUT
	A : REFERENCE TO L_UMTP_Matrix3x3;
	B : REFERENCE TO L_UMTP_Matrix3x3;
	RESULT : REFERENCE TO L_UMTP_Matrix3x3;
END_VAR
END_FUNCTION

(* ---- L_UMTP_MATRIXTIMESVECTOR3D.pou ---- *)
FUNCTION L_UMTP_MATRIXTIMESVECTOR3D
VAR_INPUT
	A : REFERENCE TO L_UMTP_Matrix3x3;
	X : REFERENCE TO L_UMTP_Vector3D;
	RESULT : REFERENCE TO L_UMTP_Vector3D;
END_VAR
END_FUNCTION

(* ---- L_UMTP_MATRIXTIMESVECTOR3DTIMESSKALAR.pou ---- *)
FUNCTION L_UMTP_MATRIXTIMESVECTOR3DTIMESSKALAR
VAR_INPUT
	A : REFERENCE TO L_UMTP_Matrix3x3;
	X : REFERENCE TO L_UMTP_Vector3D;
	SCALAR : LREAL;
	RESULT : REFERENCE TO L_UMTP_Vector3D;
END_VAR
END_FUNCTION

(* ---- L_UMTP_MATRIXTRANSPOSETIMESANTISYM3D.pou ---- *)
FUNCTION L_UMTP_MATRIXTRANSPOSETIMESANTISYM3D
VAR_INPUT
	M : REFERENCE TO L_UMTP_Matrix3x3;
	ASYM : REFERENCE TO L_UMTP_Vector3D;
	RESULT : REFERENCE TO L_UMTP_Matrix3x3;
END_VAR
END_FUNCTION

(* ---- L_UMTP_MATRIXTRANSPOSETIMESMATRIX3D.pou ---- *)
FUNCTION L_UMTP_MATRIXTRANSPOSETIMESMATRIX3D
VAR_INPUT
	A : REFERENCE TO L_UMTP_Matrix3x3;
	B : REFERENCE TO L_UMTP_Matrix3x3;
	RESULT : REFERENCE TO L_UMTP_Matrix3x3;
END_VAR
END_FUNCTION

(* ---- L_UMTP_MATRIXTRANSPOSETIMESVECTOR3D.pou ---- *)
FUNCTION L_UMTP_MATRIXTRANSPOSETIMESVECTOR3D : BOOL
VAR_INPUT
	A : REFERENCE TO L_UMTP_Matrix3x3;
	X : REFERENCE TO L_UMTP_Vector3D;
	RESULT : REFERENCE TO L_UMTP_Vector3D;
END_VAR
END_FUNCTION

(* ---- L_UMTP_MODULODIFF.pou ---- *)
FUNCTION L_UMTP_MODULODIFF : LREAL
VAR_INPUT
	LRDIFF : LREAL;
	LRCYCLELENGTH : LREAL;
	LRINVCYCLELENGTH : LREAL;
END_VAR
END_FUNCTION

(* ---- L_UMTP_MODULOPOS.pou ---- *)
FUNCTION L_UMTP_MODULOPOS : LREAL
VAR_INPUT
	LRPOSITION : LREAL;
	LRCYCLELENGTH : LREAL;
	LRINVCYCLELENGTH : LREAL;
END_VAR
VAR_OUTPUT
	LRROUNDS : LREAL;
END_VAR
END_FUNCTION

(* ---- L_UMTP_NEGMATRIX3D.pou ---- *)
FUNCTION L_UMTP_NEGMATRIX3D : BOOL
VAR_INPUT
	A : REFERENCE TO L_UMTP_Matrix3x3;
END_VAR
END_FUNCTION

(* ---- L_UMTP_NEGVECTOR3D.pou ---- *)
FUNCTION L_UMTP_NEGVECTOR3D : BOOL
VAR_INPUT
	X : REFERENCE TO L_UMTP_Vector3D;
END_VAR
END_FUNCTION

(* ---- L_UMTP_NEWTON1D.pou ---- *)
FUNCTION L_UMTP_NEWTON1D : BOOL
VAR_INPUT
	IFUNC : L_UMTP_Func_1D21D;
	CONTEXT : DINT;
	CONTEXT_DF : DINT;
	F_REQUESTED : LREAL;
	TOL : LREAL;
	X : REFERENCE TO LREAL;
END_VAR
END_FUNCTION

(* ---- L_UMTP_NORM2.pou ---- *)
FUNCTION L_UMTP_NORM2 : LREAL
VAR_INPUT
	PLRX : POINTER TO LREAL;
	UDIDIM : UDINT;
END_VAR
END_FUNCTION

(* ---- L_UMTP_NORMTO.pou ---- *)
FUNCTION L_UMTP_NORMTO : LREAL
VAR_INPUT
	PLRX : POINTER TO LREAL;
	UDIDIM : UDINT;
	VALUE : LREAL;
END_VAR
END_FUNCTION

(* ---- L_UMTP_POLY5COEFFS.pou ---- *)
FUNCTION L_UMTP_POLY5COEFFS : BOOL
VAR_INPUT
	LRY0 : LREAL;
	LRY1 : LREAL;
	LRDY0 : LREAL;
	LRDY1 : LREAL;
	LRDDY0 : LREAL;
	LRDDY1 : LREAL;
	LRL : LREAL;
END_VAR
VAR_OUTPUT
	LRA0 : LREAL;
	LRA1 : LREAL;
	LRA2 : LREAL;
	LRA3 : LREAL;
	LRA4 : LREAL;
	LRA5 : LREAL;
END_VAR
END_FUNCTION

(* ---- L_UMTP_POLYNOM.pou ---- *)
FUNCTION L_UMTP_POLYNOM : LREAL
VAR_INPUT
	PLRCOEFFS : POINTER TO LREAL;
	UDIDEGREE : UDINT;
	LRX : LREAL;
	UDIDERIV : UDINT;
END_VAR
END_FUNCTION

(* ---- L_UMTP_POLYNOMINALROOTS2.pou ---- *)
FUNCTION L_UMTP_POLYNOMINALROOTS2 : UDINT
VAR_INPUT
	FA0 : LREAL;
	FA1 : LREAL;
	FA2 : LREAL;
	LRTHRESHOLD : LREAL;
END_VAR
VAR_OUTPUT
	LRROOT0 : LREAL;
	LRROOT1 : LREAL;
END_VAR
END_FUNCTION

(* ---- L_UMTP_POLYNOMINALROOTS3.pou ---- *)
FUNCTION L_UMTP_POLYNOMINALROOTS3 : UDINT
VAR_INPUT
	PLRCOEFFS : POINTER TO LREAL;
	PLRROOTS : POINTER TO LREAL;
	LRTHRESHOLD : LREAL;
END_VAR
END_FUNCTION

(* ---- L_UMTP_POLYNOMINALROOTS4.pou ---- *)
FUNCTION L_UMTP_POLYNOMINALROOTS4 : UDINT
VAR_INPUT
	PLRCOEFFS : POINTER TO LREAL;
	PLRROOTS : POINTER TO LREAL;
	LRTHRESHOLD : LREAL;
END_VAR
END_FUNCTION

(* ---- L_UMTP_REDUCEPITCH.pou ---- *)
FUNCTION L_UMTP_REDUCEPITCH
VAR_INPUT
	FRAME : REFERENCE TO L_UMTP_RobotFrame;
	DPHIA : LREAL;
	DPHIB : LREAL;
	DPHIC : LREAL;
END_VAR
VAR_OUTPUT
	DDPHIA : LREAL;
	DDPHIB : LREAL;
	DDPHIC : LREAL;
END_VAR
END_FUNCTION

(* ---- L_UMTP_REDUCETWIST.pou ---- *)
FUNCTION L_UMTP_REDUCETWIST
VAR_INPUT
	FRAME : REFERENCE TO L_UMTP_RobotFrame;
END_VAR
VAR_OUTPUT
	DPHIA : LREAL;
	DPHIB : LREAL;
	DPHIC : LREAL;
END_VAR
END_FUNCTION

(* ---- L_UMTP_RESETROBFRAME.pou ---- *)
FUNCTION L_UMTP_RESETROBFRAME : BOOL
VAR_IN_OUT
	SCROBOTFRAME : L_UMTP_RobotFrame;
END_VAR
END_FUNCTION

(* ---- L_UMTP_RESETROBFRAMEDYNAMIC.pou ---- *)
FUNCTION L_UMTP_RESETROBFRAMEDYNAMIC : BOOL
VAR_IN_OUT
	SCROBOTFRAME : L_UMTP_RobotFrame;
END_VAR
END_FUNCTION

(* ---- L_UMTP_RESETROTMAT.pou ---- *)
FUNCTION L_UMTP_RESETROTMAT : BOOL
VAR_IN_OUT
	SCROTMAT : L_UMTP_Matrix3x3;
END_VAR
END_FUNCTION

(* ---- L_UMTP_RESOLVEGIMBALLOCKACC.pou ---- *)
FUNCTION L_UMTP_RESOLVEGIMBALLOCKACC
VAR_INPUT
	PARAM : REFERENCE TO L_UMTP_RotParam;
	DDPHIA : LREAL;
	DDPHIB : LREAL;
	DDPHIC : LREAL;
	DDPHIAOLD : LREAL;
	DDPHIBOLD : LREAL;
	DDPHICOLD : LREAL;
	T : LREAL;
	XISFIXA : BOOL;
	XISFIXB : BOOL;
	XISFIXC : BOOL;
END_VAR
VAR_OUTPUT
	DDPHIACOR : LREAL;
	DDPHIBCOR : LREAL;
	DDPHICCOR : LREAL;
END_VAR
END_FUNCTION

(* ---- L_UMTP_RESOLVEGIMBALLOCKPOS.pou ---- *)
FUNCTION L_UMTP_RESOLVEGIMBALLOCKPOS
VAR_INPUT
	PARAM : REFERENCE TO L_UMTP_RotParam;
	DPHIA : LREAL;
	DPHIB : LREAL;
	DPHIC : LREAL;
	DPHIAOLD : LREAL;
	DPHIBOLD : LREAL;
	DPHICOLD : LREAL;
	DDPHIAOLD : LREAL;
	DDPHIBOLD : LREAL;
	DDPHICOLD : LREAL;
	T : LREAL;
END_VAR
VAR_OUTPUT
	DPHIACOR : LREAL;
	DPHIBCOR : LREAL;
	DPHICCOR : LREAL;
END_VAR
END_FUNCTION

(* ---- L_UMTP_RESOLVEGIMBALLOCKVEL.pou ---- *)
FUNCTION L_UMTP_RESOLVEGIMBALLOCKVEL
VAR_INPUT
	PARAM : REFERENCE TO L_UMTP_RotParam;
	DPHIA : LREAL;
	DPHIB : LREAL;
	DPHIC : LREAL;
	DPHIAOLD : LREAL;
	DPHIBOLD : LREAL;
	DPHICOLD : LREAL;
	DDPHIAOLD : LREAL;
	DDPHIBOLD : LREAL;
	DDPHICOLD : LREAL;
	T : LREAL;
	XISFIXA : BOOL;
	XISFIXB : BOOL;
	XISFIXC : BOOL;
END_VAR
VAR_OUTPUT
	DPHIACOR : LREAL;
	DPHIBCOR : LREAL;
	DPHICCOR : LREAL;
END_VAR
END_FUNCTION

(* ---- L_UMTP_RK4STEP.pou ---- *)
FUNCTION L_UMTP_RK4STEP
VAR_INPUT
	IODE : L_UMTP_IODE;
	PLRY0 : POINTER TO LREAL;
	UDIDIM : UDINT;
	LRT : LREAL;
	LRH : LREAL;
END_VAR
VAR_OUTPUT
	LRTNEW : LREAL;
END_VAR
END_FUNCTION

(* ---- L_UMTP_ROBOTPOSTIMESFRAME.pou ---- *)
FUNCTION L_UMTP_ROBOTPOSTIMESFRAME
VAR_INPUT
	ROBOTPOS : REFERENCE TO L_UMTP_RobotPos;
	FRAME : REFERENCE TO L_UMTP_RobotFrame;
	RESULT : REFERENCE TO L_UMTP_RobotFrame;
END_VAR
END_FUNCTION

(* ---- L_UMTP_ROBOTPOSTIMESFRAMEACC.pou ---- *)
FUNCTION L_UMTP_ROBOTPOSTIMESFRAMEACC
VAR_INPUT
	ROBOTPOS : REFERENCE TO L_UMTP_RobotPos;
	FRAME : REFERENCE TO L_UMTP_RobotFrame;
	RESULT : REFERENCE TO L_UMTP_RobotFrame;
END_VAR
END_FUNCTION

(* ---- L_UMTP_ROBOTPOSTIMESFRAMEPOS.pou ---- *)
FUNCTION L_UMTP_ROBOTPOSTIMESFRAMEPOS
VAR_INPUT
	ROBOTPOS : REFERENCE TO L_UMTP_RobotPos;
	FRAME : REFERENCE TO L_UMTP_RobotFrame;
	RESULT : REFERENCE TO L_UMTP_RobotFrame;
END_VAR
END_FUNCTION

(* ---- L_UMTP_ROBOTPOSTIMESFRAMEVEL.pou ---- *)
FUNCTION L_UMTP_ROBOTPOSTIMESFRAMEVEL
VAR_INPUT
	ROBOTPOS : REFERENCE TO L_UMTP_RobotPos;
	FRAME : REFERENCE TO L_UMTP_RobotFrame;
	RESULT : REFERENCE TO L_UMTP_RobotFrame;
END_VAR
END_FUNCTION

(* ---- L_UMTP_ROBOTPOSTIMESROBOTPOS.pou ---- *)
FUNCTION L_UMTP_ROBOTPOSTIMESROBOTPOS
VAR_INPUT
	ROBOTPOSA : REFERENCE TO L_UMTP_RobotPos;
	ROBOTPOSB : REFERENCE TO L_UMTP_RobotPos;
	RESULT : REFERENCE TO L_UMTP_RobotPos;
END_VAR
END_FUNCTION

(* ---- L_UMTP_ROBOTPOSTIMESVECTOR.pou ---- *)
FUNCTION L_UMTP_ROBOTPOSTIMESVECTOR
VAR_INPUT
	ROBOTPOS : REFERENCE TO L_UMTP_RobotPos;
	A : REFERENCE TO L_UMTP_Vector3D;
	RESULT : REFERENCE TO L_UMTP_Vector3D;
END_VAR
END_FUNCTION

(* ---- L_UMTP_ROBOTPOSTOHOMMATRIX.pou ---- *)
FUNCTION L_UMTP_ROBOTPOSTOHOMMATRIX
VAR_INPUT
	HOMMATRIX : REFERENCE TO ARRAY [1..4, 1..4] OF LREAL;
	ROBOTPOS : REFERENCE TO L_UMTP_RobotPos;
	LRSCALEMATRIX2POS : LREAL;
END_VAR
END_FUNCTION

(* ---- L_UMTP_ROT2ABC.pou ---- *)
FUNCTION L_UMTP_ROT2ABC
VAR_INPUT
	ROTMAT : REFERENCE TO L_UMTP_RotMat;
	XPOSCOS2 : BOOL;
END_VAR
END_FUNCTION

(* ---- L_UMTP_ROT2QUAT.pou ---- *)
FUNCTION L_UMTP_ROT2QUAT
VAR_IN_OUT
	ROT : L_UMTP_RotMat;
	QUAT : L_UMTP_Quaternion;
END_VAR
END_FUNCTION

(* ---- L_UMTP_ROUND_LREAL.pou ---- *)
FUNCTION L_UMTP_ROUND_LREAL : LREAL
VAR_INPUT
	LRVALUE : LREAL;
END_VAR
END_FUNCTION

(* ---- L_UMTP_SCALAR.pou ---- *)
FUNCTION L_UMTP_SCALAR : LREAL
VAR_INPUT
	PLRX : POINTER TO LREAL;
	PLRY : POINTER TO LREAL;
	UDIDIM : UDINT;
END_VAR
END_FUNCTION

(* ---- L_UMTP_SCALARTIMESMATRIX3D.pou ---- *)
FUNCTION L_UMTP_SCALARTIMESMATRIX3D : BOOL
VAR_INPUT
	A : REFERENCE TO L_UMTP_Matrix3x3;
	X : LREAL;
END_VAR
END_FUNCTION

(* ---- L_UMTP_SELECTIONSORTINT.pou ---- *)
FUNCTION L_UMTP_SELECTIONSORTINT
VAR_INPUT
	PIX : POINTER TO INT;
	UDISIZE : UDINT;
	XINVERT : BOOL;
END_VAR
END_FUNCTION

(* ---- L_UMTP_SELECTIONSORTITFSORTDATA.pou ---- *)
FUNCTION L_UMTP_SELECTIONSORTITFSORTDATA : BOOL
VAR_INPUT
	ITFDATA : L_UMTP_ISortData;
	XINVERT : BOOL;
END_VAR
END_FUNCTION

(* ---- L_UMTP_SELECTIONSORTLREAL.pou ---- *)
FUNCTION L_UMTP_SELECTIONSORTLREAL
VAR_INPUT
	PLRX : POINTER TO LREAL;
	UDISIZE : UDINT;
	XINVERT : BOOL;
END_VAR
END_FUNCTION

(* ---- L_UMTP_SETIDENTITYFRAME.pou ---- *)
FUNCTION L_UMTP_SETIDENTITYFRAME
VAR_INPUT
	FRAME : REFERENCE TO L_UMTP_RobotFrame;
END_VAR
END_FUNCTION

(* ---- L_UMTP_STIMESVECTOR.pou ---- *)
FUNCTION L_UMTP_STIMESVECTOR
VAR_INPUT
	SCALAR : LREAL;
	PA : POINTER TO LREAL;
	PRESULT : POINTER TO LREAL;
	DIM : DINT;
END_VAR
END_FUNCTION

(* ---- L_UMTP_STR_IS_NUMERICALVALUE.pou ---- *)
FUNCTION L_UMTP_STR_IS_NUMERICALVALUE : BOOL
VAR_INPUT
	STVALUE : STRING(255);
END_VAR
VAR_OUTPUT
	XISINT : BOOL;
END_VAR
END_FUNCTION

(* ---- L_UMTP_STRING_TO_LREAL.pou ---- *)
FUNCTION L_UMTP_STRING_TO_LREAL : BOOL
VAR_INPUT
	STVALUE : STRING(255);
END_VAR
VAR_OUTPUT
	LRVALUE : LREAL;
END_VAR
END_FUNCTION

(* ---- L_UMTP_SWAP.pou ---- *)
FUNCTION L_UMTP_SWAP
VAR_INPUT
	A : REFERENCE TO LREAL;
	B : REFERENCE TO LREAL;
END_VAR
END_FUNCTION

(* ---- L_UMTP_THOMASALGORITHM.pou ---- *)
FUNCTION L_UMTP_THOMASALGORITHM : BOOL
VAR_INPUT
	IDIM : INT;
	ALRA : POINTER TO LREAL;
	ALRD : POINTER TO LREAL;
	ALRX : POINTER TO LREAL;
END_VAR
VAR_OUTPUT
	XERROR : BOOL := FALSE;
	EERRORID : L_IE1P_Error := L_IE1P_Error.NoError;
END_VAR
END_FUNCTION

(* ---- L_UMTP_THRESHOLD.pou ---- *)
FUNCTION L_UMTP_THRESHOLD : LREAL
VAR_INPUT
	LRVALUE : LREAL;
	LRTHRESHOLD : LREAL;
END_VAR
END_FUNCTION

(* ---- L_UMTP_TRACE.pou ---- *)
FUNCTION L_UMTP_TRACE : LREAL
VAR_IN_OUT
	ROTMAT : L_UMTP_RotMat;
END_VAR
END_FUNCTION

(* ---- L_UMTP_TRANSFERFUNCTION.pou ---- *)
FUNCTION L_UMTP_TRANSFERFUNCTION : BOOL
VAR_INPUT
	ALRIN : POINTER TO LREAL;
	ALROUT : POINTER TO LREAL;
	ALR_A : POINTER TO LREAL;
	ALR_B : POINTER TO LREAL;
END_VAR
END_FUNCTION

(* ---- L_UMTP_TRANSPOSE.pou ---- *)
FUNCTION L_UMTP_TRANSPOSE : LREAL
VAR_INPUT
	PLRM : POINTER TO LREAL;
	PLRMTRANS : POINTER TO LREAL;
	UDIROWS : UDINT;
	UDICOLS : UDINT;
END_VAR
END_FUNCTION

(* ---- L_UMTP_TRUNC_LINT.pou ---- *)
FUNCTION L_UMTP_TRUNC_LINT : LINT
VAR_INPUT
	LRIN : LREAL;
END_VAR
END_FUNCTION

(* ---- L_UMTP_VECTORADDSTIMESVECTOR.pou ---- *)
FUNCTION L_UMTP_VECTORADDSTIMESVECTOR
VAR_INPUT
	PA : POINTER TO LREAL;
	SCALAR : LREAL;
	PB : POINTER TO LREAL;
	PRESULT : POINTER TO LREAL;
	DIM : DINT;
END_VAR
END_FUNCTION

(* ---- L_UMTP_VECTORADDVECTOR.pou ---- *)
FUNCTION L_UMTP_VECTORADDVECTOR
VAR_INPUT
	PA : POINTER TO LREAL;
	PB : POINTER TO LREAL;
	PRESULT : POINTER TO LREAL;
	DIM : DINT;
END_VAR
END_FUNCTION

(* ---- L_UMTP_VECTORANGLE3D.pou ---- *)
FUNCTION L_UMTP_VECTORANGLE3D : BOOL
VAR_INPUT
	A : REFERENCE TO ARRAY [1..3] OF LREAL;
	B : REFERENCE TO ARRAY [1..3] OF LREAL;
	RESULT : REFERENCE TO LREAL;
END_VAR
END_FUNCTION

(* ---- L_UMTP_VECTORCOLLINEAR3D.pou ---- *)
FUNCTION L_UMTP_VECTORCOLLINEAR3D : BOOL
VAR_INPUT
	A : REFERENCE TO ARRAY [1..3] OF LREAL;
	B : REFERENCE TO ARRAY [1..3] OF LREAL;
END_VAR
END_FUNCTION

(* ---- L_UMTP_VECTOREQUALS.pou ---- *)
FUNCTION L_UMTP_VECTOREQUALS : BOOL
VAR_INPUT
	PV0 : POINTER TO LREAL;
	PV1 : POINTER TO LREAL;
	ICOUNT : INT;
END_VAR
END_FUNCTION

(* ---- L_UMTP_VECTORTHRESHOLD.pou ---- *)
FUNCTION L_UMTP_VECTORTHRESHOLD
VAR_INPUT
	PLRVALUE : POINTER TO LREAL;
	UDIDIM : UDINT;
	LRTHRESHOLD : LREAL;
END_VAR
END_FUNCTION

(* ---- L_UMTP_WRITEMATRIXTOFILE.pou ---- *)
FUNCTION L_UMTP_WRITEMATRIXTOFILE : BOOL
VAR_INPUT
	PLRMAT : POINTER TO LREAL;
	UDIROWS : UDINT;
	UDICOLS : UDINT;
	FILENAME : STRING;
END_VAR
END_FUNCTION

(* ---- L_UMTP_WRITEPATHTOFILE.pou ---- *)
FUNCTION L_UMTP_WRITEPATHTOFILE : BOOL
VAR_INPUT
	IPATH : L_UMTP_IPath;
	N : UDINT;
	XWRITEPOS : BOOL;
	XWRITED1 : BOOL;
	XWRITED2 : BOOL;
	FILENAME : STRING;
END_VAR
END_FUNCTION

(* ---- REPLACE_WITH.pou ---- *)
FUNCTION REPLACE_WITH : STRING(255)
VAR_INPUT
	STR : STRING(255);
	OLD : STRING(255);
	NEW : STRING(255);
END_VAR
END_FUNCTION

(* ---- GLOBALTEXTLIST.pou ---- *)
FUNCTION_BLOCK GLOBALTEXTLIST
VAR
	M_TEXTLISTFILE : STRING(255);
	_STNAMESPACE : STRING;
END_VAR
END_FUNCTION_BLOCK

(* ---- L_UMTP_2DINTERPOLATION.pou ---- *)
FUNCTION_BLOCK L_UMTP_2DINTERPOLATION
VAR_INPUT
	XENABLE : BOOL;
	ALRX : POINTER TO LREAL;
	DINBROFXVALUES : DINT := -1;
	EINTERPTYPEX : L_UMTP_InterpolationType := L_UMTP_InterpolationType.Linear;
	ALRY : POINTER TO LREAL;
	DINBROFYVALUES : DINT := -1;
	EINTERPTYPEY : L_UMTP_InterpolationType := L_UMTP_InterpolationType.Linear;
	ALRZ : POINTER TO LREAL;
	LRX : LREAL;
	LRY : LREAL;
END_VAR
VAR_OUTPUT
	XVALID : BOOL;
	XERROR : BOOL;
	EERRORID : L_IE1P_Error;
	LRZ : LREAL;
END_VAR
VAR
	LININTERP : L_UMTP_InterpolationLinear;
	SPLINEINTERP : L_UMTP_InterpolationCubicSpline;
	INTERPDATA : L_UMTP_InterpolationData;
	ALRZROW_FOR_ALRY : ARRAY [1..cdiMaxValuesX] OF LREAL;
	ALRINTERPZCOL_AT_LRX : ARRAY [1..cdiMaxValuesY] OF LREAL;
	IDX1 : DINT;
	IDX2 : DINT;
	LRXOLD : LREAL := L_UMTP_Math.L_UMTP_ValueInitial;
	LRX_INT : LREAL;
	LRY_INT : LREAL;
	DINBROFXVALUES_INT : DINT;
	DINBROFYVALUES_INT : DINT;
	XENABLEOLD : BOOL;
	CDIMAXVALUESX : DINT := 10;
	CDIMAXVALUESY : DINT := 10;
END_VAR
END_FUNCTION_BLOCK

(* ---- L_UMTP_CALCMONOTONRISINGROTVEC.pou ---- *)
FUNCTION_BLOCK L_UMTP_CALCMONOTONRISINGROTVEC
VAR
	SCVECTORDIRECTIONINIT : L_UMTP_Vector3D;
	LRVECTORNORMINTE : LREAL := 0.0;
	LRVECTORNORMOLD : LREAL := 0.0;
	LRVECTORLENGTH : LREAL;
END_VAR
END_FUNCTION_BLOCK

METHOD CALCROTVEC : BOOL
VAR_OUTPUT
	SCROTVECTOR : L_UMTP_Vector3D;
END_VAR
VAR_IN_OUT
	SCACTROTMATRIX : L_UMTP_RotMat;
END_VAR
END_METHOD

METHOD INIT : BOOL
VAR_IN_OUT
	SCINITROTMATRIX : L_UMTP_RotMat;
END_VAR
END_METHOD

METHOD RESET : BOOL
END_METHOD

(* ---- L_UMTP_COXDEBOORCOEFFICIENTS.pou ---- *)
FUNCTION_BLOCK L_UMTP_COXDEBOORCOEFFICIENTS
VAR_INPUT
	LRU : LREAL;
	UDITODEGREE : UDINT;
	UDIINTERVAL : REFERENCE TO UDINT;
END_VAR
VAR_OUTPUT
	XERROR : BOOL;
END_VAR
VAR
	M_ALRKNOTS : ARRAY [0..(udiMaxm_alrKnots - 1)] OF LREAL;
	M_ALRNIJ : ARRAY [0..(udiMaxm_alrKnots - 1)] OF LREAL;
	M_NKNOTS : UDINT;
	Z : LREAL;
	N : LREAL;
	M_ACTDEGREE : UDINT;
	M_DEGREE : UDINT;
	I : UDINT;
	D : UDINT;
	UDIMAXM_ALRKNOTS : UDINT := 100;
	KNOTS : POINTER TO LREAL;
	NIJ : POINTER TO LREAL;
END_VAR
END_FUNCTION_BLOCK

METHOD FINDINTERVALINTERNAL : BOOL
VAR_INPUT
	LRU : LREAL;
	UDIINTERVAL : REFERENCE TO UDINT;
END_VAR
END_METHOD

METHOD PREPAREUNIFORM : BOOL
VAR_INPUT
	UDINCP : UDINT;
	UDIDEGREE : UDINT;
END_VAR
END_METHOD

METHOD PREPAREWITH : BOOL
VAR_INPUT
	ALRU : POINTER TO LREAL;
END_VAR
END_METHOD

METHOD RESET
END_METHOD

(* ---- L_UMTP_ENSURESTEADY.pou ---- *)
FUNCTION_BLOCK L_UMTP_ENSURESTEADY
VAR_INPUT
	XENABLE : BOOL;
	LRINPUT : LREAL;
	LRINPUTVELMAX : LREAL;
	LRCYCLE : LREAL;
END_VAR
VAR_OUTPUT
	XISSTEADY : BOOL := TRUE;
END_VAR
VAR
	XENABLE_OLD : BOOL := FALSE;
	LRINPUT_OLD : LREAL;
	LRINPUTVEL : LREAL;
END_VAR
END_FUNCTION_BLOCK

(* ---- L_UMTP_FFTDATA.pou ---- *)
FUNCTION_BLOCK L_UMTP_FFTDATA
VAR
	_PLCINPUTDATA : POINTER TO L_UMTP_Complex;
	_PLCOUTPUTDATA : POINTER TO L_UMTP_Complex;
	_UDIDATACOUNT : UDINT;
	_UDIARRAYLENGTH : UDINT;
	_XERROR : BOOL;
	_RESOURCEHANDLING : L_UBUP_criticalsection;
	_XLOCKED : BOOL;
	_DWITERCURRENT : DWORD;
	CURRENT : DWORD;
	HASNEXT : BOOL;
	HASPREV : BOOL;
	ITFITERATOR : L_UBUP.L_UBUP_IIterator;
	ITFLISTCONTROL : L_UBUP_IListControl;
	LENGTH : UDINT;
	PTRINPUTDATA : POINTER TO L_UMTP_Complex;
	PTROUTPUTDATA : POINTER TO L_UMTP_Complex;
END_VAR
END_FUNCTION_BLOCK

METHOD NEXT : DWORD
END_METHOD

METHOD PREV : DWORD
END_METHOD

METHOD REWIND
VAR_OUTPUT
	DWARRAYIDXSTART : DWORD;
END_VAR
END_METHOD

METHOD LOCK : BOOL
END_METHOD

METHOD LOCKSTATE : BOOL
END_METHOD

METHOD UNLOCK : BOOL
END_METHOD

METHOD GETSTRING : BOOL
VAR_INPUT
	DWARRIDX : DWORD;
END_VAR
VAR_OUTPUT
	STVALUE : STRING(255);
END_VAR
END_METHOD

METHOD REQUESTINTERFACE : BOOL
VAR_INPUT
	ID : DINT;
	PITFUNKNOWN : POINTER TO L_UBUP_IUnknown;
END_VAR
END_METHOD

METHOD RECORDDATA : UDINT
VAR_INPUT
	PLCDATA : POINTER TO L_UMTP_Complex;
	UDISIZEOFDATA : UDINT;
END_VAR
END_METHOD

METHOD STARTRECORDING : BOOL
END_METHOD

METHOD STOPRECORDING : BOOL
END_METHOD

METHOD FB_INIT : BOOL
VAR_INPUT
	BINITRETAINS : BOOL;
	BINCOPYCODE : BOOL;
END_VAR
END_METHOD

(* ---- L_UMTP_FFTDATA2048.pou ---- *)
FUNCTION_BLOCK L_UMTP_FFTDATA2048 EXTENDS L_UMTP_FFTData
VAR
	ALCDATAIN : ARRAY [1..c_arraylength] OF L_UMTP_Complex;
	ALCDATAOUT : ARRAY [1..c_arraylength] OF L_UMTP_Complex;
	C_ARRAYLENGTH : UDINT := 2048;
END_VAR
END_FUNCTION_BLOCK

METHOD GETSTRING : BOOL
VAR_INPUT
	DWARRIDX : DWORD;
END_VAR
VAR_OUTPUT
	STVALUE : STRING(255);
END_VAR
END_METHOD

METHOD FB_INIT : BOOL
VAR_INPUT
	BINITRETAINS : BOOL;
	BINCOPYCODE : BOOL;
END_VAR
END_METHOD

METHOD FB_REINIT : BOOL
END_METHOD

(* ---- L_UMTP_GOODNESSOFFIT.pou ---- *)
FUNCTION_BLOCK L_UMTP_GOODNESSOFFIT
VAR_INPUT
	XENABLE : BOOL;
	LRX : LREAL;
	LRXREF : LREAL;
	LRLAMBDA : LREAL := 1.0;
END_VAR
VAR_OUTPUT
	LRNRMSE : LREAL;
	LRNMSE : LREAL;
END_VAR
VAR
	LRSUMOFX : LREAL;
	LRSUMOFXSQR : LREAL;
	LRNUMERATOR : LREAL;
	LRDENOMINATOR : LREAL;
	LRINVDENOMINATOR : LREAL;
	LRNBROFCYCLES : LREAL;
END_VAR
END_FUNCTION_BLOCK

(* ---- L_UMTP_HYSTERESIS.pou ---- *)
FUNCTION_BLOCK L_UMTP_HYSTERESIS
VAR_INPUT
	LRIN : LREAL;
	LRHYSTERESISWIDTH : LREAL := 0;
END_VAR
VAR_OUTPUT
	XBUSY : BOOL;
	XERROR : BOOL;
	EERRORID : L_IE1P_Error;
	LROUT : LREAL;
END_VAR
VAR
	LROUT_OLD : LREAL := 0;
	LROLDHYSTWIDTH : LREAL;
	ISTEP : INT := 0;
END_VAR
END_FUNCTION_BLOCK

(* ---- L_UMTP_INTERPOLATIONBASE.pou ---- *)
FUNCTION_BLOCK L_UMTP_INTERPOLATIONBASE
VAR_INPUT
	SCDATA : L_UMTP_InterpolationData;
END_VAR
VAR_OUTPUT
	XISREADY : BOOL;
	XERROR : BOOL;
	EERRORID : L_IE1P_Error;
END_VAR
VAR
	XTRYFIRST : BOOL;
	UDNINTERVAL : UDINT;
	LRDX : LREAL;
	LRDY : LREAL;
	INTERPOLATIONTYPE : L_UMTP_InterpolationType;
	XMAX : LREAL;
	XMIN : LREAL;
END_VAR
END_FUNCTION_BLOCK

METHOD CHECKFORSTRICTLYMONOTONIC : BOOL
END_METHOD

METHOD GETVALUE : BOOL
VAR_INPUT
	X : LREAL;
END_VAR
VAR_OUTPUT
	Y : LREAL;
END_VAR
END_METHOD

METHOD GETVALUEIMPL : BOOL
VAR_INPUT
	X : LREAL;
END_VAR
VAR_OUTPUT
	Y : LREAL;
END_VAR
END_METHOD

METHOD GET_XI : LREAL
VAR_INPUT
	IDX : UDINT;
END_VAR
END_METHOD

METHOD GET_YI : LREAL
VAR_INPUT
	IDX : UDINT;
END_VAR
END_METHOD

METHOD WRITETOFILE : BOOL
VAR_INPUT
	PATH : STRING;
END_VAR
END_METHOD

(* ---- L_UMTP_INTERPOLATIONCUBICSPLINE.pou ---- *)
FUNCTION_BLOCK L_UMTP_INTERPOLATIONCUBICSPLINE EXTENDS L_UMTP_InterpolationBase
VAR_INPUT
	EINTERPOLATIONTYPE : L_UMTP_InterpolationType := L_UMTP_InterpolationType.CubicSplineHermite;
	LRSLOPE0 : LREAL;
	LRSLOPEN : LREAL;
END_VAR
VAR
	ALRSPLINECOEFFS : ARRAY [0..(L_UMTP_Constants.gc_udiMaxCubSplinePts - 2)] OF ARRAY [1..4] OF LREAL;
	ALRH : ARRAY [0..(L_UMTP_Constants.gc_udiMaxCubSplinePts - 2)] OF LREAL;
	ALRINVH : ARRAY [0..(L_UMTP_Constants.gc_udiMaxCubSplinePts - 2)] OF LREAL;
	ALRX : ARRAY [0..(L_UMTP_Constants.gc_udiMaxCubSplinePts - 1), 1..1] OF LREAL;
	ALRA : ARRAY [0..(L_UMTP_Constants.gc_udiMaxCubSplinePts - 1), 1..3] OF LREAL;
	ALRD : ARRAY [0..(L_UMTP_Constants.gc_udiMaxCubSplinePts - 1), 1..1] OF LREAL;
	EINTERPOLATIONTYPEINT : L_UMTP_InterpolationType;
	INTERPOLATIONTYPE : L_UMTP_InterpolationType;
END_VAR
END_FUNCTION_BLOCK

METHOD CALCSPLINECOEFF : BOOL
END_METHOD

METHOD GETVALUEIMPL : BOOL
VAR_INPUT
	X : LREAL;
END_VAR
VAR_OUTPUT
	Y : LREAL;
END_VAR
END_METHOD

(* ---- L_UMTP_INTERPOLATIONLINEAR.pou ---- *)
FUNCTION_BLOCK L_UMTP_INTERPOLATIONLINEAR EXTENDS L_UMTP_InterpolationBase
VAR
	INTERPOLATIONTYPE : L_UMTP_InterpolationType;
END_VAR
END_FUNCTION_BLOCK

METHOD GETVALUEIMPL : BOOL
VAR_INPUT
	X : LREAL;
END_VAR
VAR_OUTPUT
	Y : LREAL;
END_VAR
END_METHOD

(* ---- L_UMTP_INTERPOLATIONNEWTON.pou ---- *)
FUNCTION_BLOCK L_UMTP_INTERPOLATIONNEWTON EXTENDS L_UMTP_InterpolationBase
VAR
	INTERPOLATIONTYPE : L_UMTP_InterpolationType;
END_VAR
END_FUNCTION_BLOCK

METHOD GETVALUEIMPL : BOOL
VAR_INPUT
	X : LREAL;
END_VAR
VAR_OUTPUT
	Y : LREAL;
END_VAR
END_METHOD

(* ---- L_UMTP_NUMDIFFROBFRAME.pou ---- *)
FUNCTION_BLOCK L_UMTP_NUMDIFFROBFRAME
VAR
	SCPOSVECTORMINUS0 : L_UMTP_Vector3D;
	SCPOSVECTORMINUS1 : L_UMTP_Vector3D;
	SCPOSVECTORMINUS2 : L_UMTP_Vector3D;
	SCROTMINUS0 : L_UMTP_Matrix3x3;
	SCROTMINUS1 : L_UMTP_Matrix3x3;
	SCROTMINUS2 : L_UMTP_Matrix3x3;
	XUSEROTVEC : BOOL := FALSE;
	ICNTCYCLES : INT;
	SCTWISTSTART : L_UMTP_Vector3D;
	SCPITCHSTART : L_UMTP_Vector3D;
	SCVELSTART : L_UMTP_Vector3D;
	SCACCSTART : L_UMTP_Vector3D;
END_VAR
END_FUNCTION_BLOCK

METHOD INIT : BOOL
VAR_IN_OUT
	SCFRAME : L_UMTP_RobotFrame;
END_VAR
END_METHOD

METHOD NUMDIFF : BOOL
VAR_INPUT
	LRTIMEINV : LREAL;
END_VAR
VAR_IN_OUT
	SCFRAME : L_UMTP_RobotFrame;
END_VAR
END_METHOD

METHOD RESET : BOOL
END_METHOD

METHOD UPDATEFRAMEDATAS : BOOL
VAR_IN_OUT
	SCFRAME : L_UMTP_RobotFrame;
END_VAR
END_METHOD

(* ---- L_UMTP_NUMERCALJACOBI.pou ---- *)
FUNCTION_BLOCK L_UMTP_NUMERCALJACOBI
VAR_INPUT
	IFUNC : L_UMTP_Func_ND2MD;
	CONTEXT : UDINT;
	UDIXDIM : UDINT;
	UDIYDIM : UDINT;
	ALRAT : ARRAY [1..10] OF LREAL;
END_VAR
VAR
	ALRMAT : ARRAY [1..(10 * 10)] OF LREAL;
	I : UDINT;
	J : UDINT;
	ALRPOS : ARRAY [1..10] OF LREAL;
	ALRYFWD : ARRAY [1..10] OF LREAL;
	ALRYBWD : ARRAY [1..10] OF LREAL;
	H : LREAL := 1E-06;
	COLS : UDINT;
	PTR : POINTER TO LREAL;
	ROWS : UDINT;
END_VAR
END_FUNCTION_BLOCK

METHOD GETVALUE : LREAL
VAR_INPUT
	I : UDINT;
	J : UDINT;
END_VAR
END_METHOD

METHOD SETVALUE
VAR_INPUT
	I : UDINT;
	J : UDINT;
	VALUE : LREAL;
END_VAR
END_METHOD

(* ---- L_UMTP_PATHBSPLINE.pou ---- *)
FUNCTION_BLOCK L_UMTP_PATHBSPLINE
VAR_INPUT
	PLRCP : POINTER TO LREAL;
	UDINCP : UDINT;
	UDIDIM : UDINT;
	UDIDEGREE : UDINT;
	XINITUNIFORMKNOTS : BOOL;
END_VAR
VAR_OUTPUT
	XREADY : BOOL;
	XERROR : BOOL;
END_VAR
VAR
	M_UDIDIM : UDINT;
	M_UDIDEGREE : UDINT;
	M_UDINCP : UDINT;
	M_FBCOXDEBOOR : L_UMTP_CoxdeBoorCoefficients;
	COXDEBOOR : REFERENCE TO L_UMTP_CoxdeBoorCoefficients;
	DIM : UDINT;
END_VAR
END_FUNCTION_BLOCK

METHOD GETPATHVALUE : BOOL
VAR_INPUT
	PLRX : POINTER TO LREAL;
	PLRD1 : POINTER TO LREAL;
	PLRD2 : POINTER TO LREAL;
	UDIDIM : UDINT;
	LRU : LREAL;
END_VAR
END_METHOD

(* ---- L_UMTP_PATHNURBS.pou ---- *)
FUNCTION_BLOCK L_UMTP_PATHNURBS EXTENDS L_UMTP_PathBSpline
VAR_INPUT
	PLRWEIGHTS : POINTER TO LREAL;
END_VAR
VAR
	M_PLRWEIGHTS : POINTER TO LREAL;
END_VAR
END_FUNCTION_BLOCK

METHOD GETPATHVALUE : BOOL
VAR_INPUT
	PLRX : POINTER TO LREAL;
	PLRD1 : POINTER TO LREAL;
	PLRD2 : POINTER TO LREAL;
	UDIDIM : UDINT;
	LRU : LREAL;
END_VAR
END_METHOD

(* ---- L_UMTP_PATHPOLY5.pou ---- *)
FUNCTION_BLOCK L_UMTP_PATHPOLY5
VAR_INPUT
	PLRY0 : POINTER TO LREAL;
	PLRDY0 : POINTER TO LREAL;
	PLRDDY0 : POINTER TO LREAL;
	PLRY1 : POINTER TO LREAL;
	PLRDY1 : POINTER TO LREAL;
	PLRDDY1 : POINTER TO LREAL;
	UDIDIM : UDINT;
END_VAR
VAR_OUTPUT
	XREADY : BOOL;
	XERROR : BOOL;
END_VAR
VAR
	M_ALRCOEFFS : ARRAY [1..8, 1..6] OF LREAL;
	M_UDIDIM : UDINT;
	DIM : UDINT;
END_VAR
END_FUNCTION_BLOCK

METHOD GETPATHVALUE : BOOL
VAR_INPUT
	PLRX : POINTER TO LREAL;
	PLRD1 : POINTER TO LREAL;
	PLRD2 : POINTER TO LREAL;
	UDIDIM : UDINT;
	LRU : LREAL;
END_VAR
END_METHOD

(* ---- L_UMTP_PENTADIAGONALSOLVER.pou ---- *)
FUNCTION_BLOCK L_UMTP_PENTADIAGONALSOLVER
VAR_INPUT
	PLRCHASINGPOINTS : POINTER TO LREAL;
	UDINCP : UDINT;
	UDIDIM : UDINT;
	COXDEBOOR : REFERENCE TO L_UMTP_CoxdeBoorCoefficients;
END_VAR
VAR_OUTPUT
	X : ARRAY [1..(L_UMTP_Constants.gc_iMaxNumOfGivenPts + 1), 1..3] OF LREAL;
	U : ARRAY [1..L_UMTP_Constants.gc_CtrlPtMaxNr] OF LREAL;
	V : ARRAY [1..L_UMTP_Constants.gc_CtrlPtMaxNr] OF LREAL;
END_VAR
VAR
	UDIDEGREE : DINT := 3;
	A : ARRAY [1..(L_UMTP_Constants.gc_iMaxNumOfGivenPts + 1), 1..(L_UMTP_Constants.gc_iMaxNumOfGivenPts + 1)] OF LREAL;
	B : ARRAY [1..(L_UMTP_Constants.gc_iMaxNumOfGivenPts + 1), 1..3] OF LREAL;
	D : ARRAY [1..(L_UMTP_Constants.gc_iMaxNumOfGivenPts + 1)] OF LREAL;
	E : ARRAY [1..(L_UMTP_Constants.gc_iMaxNumOfGivenPts + 1)] OF LREAL;
	F : ARRAY [1..(L_UMTP_Constants.gc_iMaxNumOfGivenPts + 1)] OF LREAL;
	G : ARRAY [1..(L_UMTP_Constants.gc_iMaxNumOfGivenPts + 1)] OF LREAL;
	H : ARRAY [1..(L_UMTP_Constants.gc_iMaxNumOfGivenPts + 1)] OF LREAL;
	ALPHA : ARRAY [1..(L_UMTP_Constants.gc_iMaxNumOfGivenPts + 1)] OF LREAL;
	DELTA : ARRAY [1..(L_UMTP_Constants.gc_iMaxNumOfGivenPts + 1)] OF LREAL;
	C : ARRAY [1..(L_UMTP_Constants.gc_iMaxNumOfGivenPts + 1), 1..3] OF LREAL;
	BET : ARRAY [1..(L_UMTP_Constants.gc_iMaxNumOfGivenPts + 1)] OF LREAL;
	GAM : ARRAY [1..(L_UMTP_Constants.gc_iMaxNumOfGivenPts + 1)] OF LREAL;
	I : INT;
	J : INT;
	K : INT;
	N : INT;
	STSTARTTIME : SysTime;
	STENDTIME : SysTime;
	STCALCULATETIME : SysTime;
	MATRIXTEST : ARRAY [1..7, 1..7] OF LREAL;
END_VAR
END_FUNCTION_BLOCK

METHOD CODEVONWERNI
END_METHOD

(* ---- L_UMTP_RADIX2FFT.pou ---- *)
FUNCTION_BLOCK L_UMTP_RADIX2FFT EXTENDS L_UBUP_FreeRunTask
VAR_INPUT
	ITFFFTDATA : L_UMTP_IFFTData;
	XIFFT : BOOL;
END_VAR
VAR_OUTPUT
	XACTIVE : BOOL := FALSE;
END_VAR
VAR
	_ITFRESOURCEHANDLING : L_UBUP_ILockable;
	_XLOCK : BOOL;
END_VAR
END_FUNCTION_BLOCK

METHOD EXECUTEIMPL : UDINT
END_METHOD

METHOD FINALIZEACTION
VAR_INPUT
	XABORTPROPOSED : BOOL;
	IERRORIDPROPOSED : INT;
END_VAR
VAR_OUTPUT
	XCOMPLETE : BOOL;
	XABORT : BOOL;
	IERRORID : INT;
END_VAR
END_METHOD

METHOD STARTACTION
VAR_OUTPUT
	XCOMPLETE : BOOL;
	IERRORID : INT;
END_VAR
END_METHOD

METHOD FFT_RADIX2 : BOOL
VAR_INPUT
	P_X : POINTER TO L_UMTP_Complex;
	UDISIZE : UDINT;
END_VAR
END_METHOD

(* ---- L_UMTP_RANDOMGENERATOR.pou ---- *)
FUNCTION_BLOCK L_UMTP_RANDOMGENERATOR
VAR_INPUT
	XENABLE : BOOL;
	LRMAXVALUE : LREAL := 1;
	LRMINVALUE : LREAL := 0;
	DWIDX : DWORD := 1;
	WRANDOMMODE : WORD := 0;
	DWSEEDVALUETOSET : DWORD := 0;
END_VAR
VAR_OUTPUT
	ALRRESULT : ARRAY [1..dwMaxRndResults] OF LREAL;
	XERROR : BOOL := FALSE;
	SERRMSG : STRING;
	DWSEEDVALUE : DWORD;
END_VAR
VAR
	DWACTRANDOMVALUE : DWORD;
	DWACTRANDOMVALUE2 : DWORD;
	LRACTRANDOMVALUE : LREAL;
	LRACTRANDOMVALUE2 : LREAL;
	DWFIRSTVALUE : DWORD := 0;
	DWFACTOR : DWORD := 65;
	DWCTR : DWORD;
	DWCTR1 : DWORD;
	XENABLEOLD : BOOL;
	LRTEMPVAR : LREAL;
	LRVARIANCE : LREAL;
	LRSIGMA : LREAL;
	LRMU : LREAL;
	DWMAXRNDRESULTS : DWORD := 255;
	DWINKREMENT : DWORD := 1;
	DWMODULO : DWORD := 99971;
	LRINVMODULO : LREAL := (1 / DWORD_TO_LREAL(dwModulo));
END_VAR
END_FUNCTION_BLOCK

(* ---- L_UMTP_RLS.pou ---- *)
FUNCTION_BLOCK L_UMTP_RLS
VAR_INPUT
	XENABLE : BOOL;
	WMODE : WORD;
	LRLAMBDA : LREAL := 1;
	PLRYK : POINTER TO LREAL;
	PLRPSIK : POINTER TO LREAL;
	PLRPARAMIN : POINTER TO LREAL;
	PLRPARAMAX : POINTER TO LREAL;
	PLRPARAK : POINTER TO LREAL;
	USIDIMY : USINT;
	USIDIMPARA : USINT;
	AUSIDIMPSI : ARRAY [1..2] OF USINT;
END_VAR
VAR_OUTPUT
	XERROR : BOOL;
END_VAR
VAR
	LRYKI : LREAL;
	ALRPK : ARRAY [1..cusiMaxPar, 1..cusiMaxPar] OF LREAL;
	ALRLK : ARRAY [1..cusiMaxPar] OF LREAL;
	ALRPK_PSIKI : ARRAY [1..cusiMaxPar] OF LREAL;
	ALRPSIKIT_PK : ARRAY [1..cusiMaxPar] OF LREAL;
	LRPSIKIT_PK_PSIKI : LREAL;
	LRPSIKIT_PARA : LREAL;
	LRDEVIATION : LREAL;
	PLRPSIKI : POINTER TO LREAL;
	ALRPSIKI : ARRAY [1..cusiMaxPar] OF LREAL;
	XENABLEOLD : BOOL;
	IDXPARROWS : USINT;
	IDXPARCOLUMNS : USINT;
	IDXMEASURE : USINT;
	LRLAMBDAINT : LREAL;
	USIDIMYINT : USINT;
	USIDIMPARAINT : USINT;
	AUSIDIMPSIINT : ARRAY [1..2] OF USINT;
	LRINVLAMBDA : LREAL;
	LRNENNER : LREAL;
	LRINVNENNER : LREAL;
	PLRTEMP : POINTER TO LREAL;
	PLRTEMP2 : POINTER TO LREAL;
	LRTEMP : LREAL;
	LRTEMP2 : LREAL;
	XINIT : BOOL := FALSE;
	XNEWPARINSIDELIMITS : BOOL;
	ALRMINSENSITIVITY : ARRAY [1..cusiMaxPar] OF LREAL;
	ALRMAXSENSITIVITY : ARRAY [1..cusiMaxPar] OF LREAL;
	XSENSITIVITYAVAILABLE : BOOL;
	LRACTABSSENSITIVITY : LREAL;
	LRSENSITIVITYTOL1 : LREAL := 0.01;
	LRSENSITIVITYTOL2 : LREAL := 0.15;
	CUSIMAXPAR : USINT := 30;
	CUSIMAXMEASURE : USINT := 6;
END_VAR
END_FUNCTION_BLOCK

(* ---- L_UMTP_SHUNTINGYARDALGORITHM.pou ---- *)
FUNCTION_BLOCK L_UMTP_SHUNTINGYARDALGORITHM
VAR_INPUT
	SINPUT : STRING(255);
	ETRIGUNIT : L_UMTP_TrigonometricUnit := L_UMTP_TrigonometricUnit.Radiant;
END_VAR
VAR_OUTPUT
	SCVALUE : L_UBUP_Variable;
	XVALID : BOOL;
	XERROR : BOOL;
	EERRORID : L_IE1P_Error := L_IE1P_Error.NoError;
END_VAR
VAR
	AEREVERSEPOLISHNOTATIONVARVALUE : ARRAY [1..255] OF L_UBUP_VarValue;
	AEREVERSEPOLISHNOTATIONOPERATOR : ARRAY [1..255] OF L_UMTP_ReversePolishNotationToken;
	INUMBEROFENTRIES : UDINT;
	AOPERATORSTACK : ARRAY [1..255] OF L_UMTP_ReversePolishNotationToken;
	ISTACKCOUNTER : UDINT;
	_SSTRING : STRING(255);
	CINBROFTOKENS : INT := 38;
END_VAR
END_FUNCTION_BLOCK

METHOD CALL_FBMETHODS
END_METHOD

METHOD CALL_OUTPUT
END_METHOD

METHOD CALL_RESETOUTPUTS
END_METHOD

METHOD FUN_COMPAREPRECEDENCE : BOOL
VAR_INPUT
	TOKEN1 : L_UMTP_ReversePolishNotationToken;
	TOKEN2 : L_UMTP_ReversePolishNotationToken;
END_VAR
END_METHOD

METHOD FUN_EVALUATEREVERSEPOLISHNOTATION : BOOL
VAR_OUTPUT
	SCVALUE : L_UBUP_Variable;
	XERROR : BOOL := FALSE;
	EERRORID : L_IE1P_Error := 0;
END_VAR
END_METHOD

METHOD FUN_ISOPERATOR : BOOL
VAR_INPUT
	TOKEN : L_UMTP_ReversePolishNotationToken;
END_VAR
END_METHOD

METHOD FUN_NEXTTOKEN : BOOL
VAR_OUTPUT
	TOKEN : STRING;
END_VAR
VAR_IN_OUT
	STR : STRING(255);
END_VAR
END_METHOD

METHOD FUN_POPSTACKIF
VAR_INPUT
	TOKEN : L_UMTP_ReversePolishNotationToken;
END_VAR
END_METHOD

METHOD FUN_PREPARELINE
VAR_IN_OUT
	SSTRING : STRING(255);
END_VAR
END_METHOD

METHOD FUN_SHUNTING_YARD_ALGORITHM : BOOL
VAR_OUTPUT
	XERROR : BOOL;
	EERRORID : L_IE1P_Error;
END_VAR
VAR_IN_OUT
	STR : STRING(255);
END_VAR
END_METHOD

METHOD FUN_TOKENPRIORITY : BOOL
VAR_INPUT
	TOKEN : L_UMTP_ReversePolishNotationToken;
END_VAR
VAR_OUTPUT
	UIPRIORITY : UINT;
END_VAR
END_METHOD

(* ---- L_UMTP_SOLVE_EQUATIONS_CHASINGMETHOD.pou ---- *)
FUNCTION_BLOCK L_UMTP_SOLVE_EQUATIONS_CHASINGMETHOD
VAR_INPUT
	Q : POINTER TO LREAL;
	COXDEBOOR : REFERENCE TO L_UMTP_CoxdeBoorCoefficients;
END_VAR
VAR_OUTPUT
	CONTRO_POS : ARRAY [1..3, 1..L_UMTP_Constants.gc_CtrlPtMaxNr] OF LREAL;
END_VAR
VAR
	N : INT;
	M : ARRAY [1..L_UMTP_Constants.gc_CtrlPtMaxNr, 1..L_UMTP_Constants.gc_CtrlPtMaxNr] OF LREAL;
	I : INT;
	J : INT;
	D : ARRAY [1..L_UMTP_Constants.gc_CtrlPtMaxNr] OF LREAL;
	U : ARRAY [1..L_UMTP_Constants.gc_CtrlPtMaxNr] OF LREAL;
	L : ARRAY [1..L_UMTP_Constants.gc_CtrlPtMaxNr] OF LREAL;
	B : ARRAY [1..L_UMTP_Constants.gc_CtrlPtMaxNr] OF LREAL;
END_VAR
END_FUNCTION_BLOCK

(* ---- L_UMTP_STATISTICS.pou ---- *)
FUNCTION_BLOCK L_UMTP_STATISTICS
VAR_INPUT
	XENABLE : BOOL;
	LRINPUT : LREAL;
END_VAR
VAR_OUTPUT
	XBUSY : BOOL;
	LRAVERAGE : LREAL;
	LRVARIANCE : LREAL;
	LRSTANDARDDEVIATION : LREAL;
	LRMIN : LREAL;
	LRMAX : LREAL;
	XOVERRUN : BOOL;
END_VAR
VAR
	LRCOUNTER : LREAL;
	LRAVERAGEINTERNAL : LREAL;
	LRVARIANCEINTERNAL : LREAL;
	LRVARIANCEINTERNAL2 : LREAL;
	LRAVERAGEOLD : LREAL;
	XENABLEOLD : BOOL;
	LRMINVALUEINT : LREAL;
	LRMAXVALUEINT : LREAL;
END_VAR
END_FUNCTION_BLOCK

(* ---- L_UMTP_TRACEFFTDATA.pou ---- *)
FUNCTION_BLOCK L_UMTP_TRACEFFTDATA
VAR_INPUT
	ITFFFTDATA : L_UMTP_IFFTData;
	XEXECUTE : BOOL;
	XABORT : BOOL;
END_VAR
VAR_OUTPUT
	XDONE : BOOL;
	XBUSY : BOOL;
	XACTIVE : BOOL;
	XCOMMANDABORTED : BOOL;
	XERROR : BOOL;
	EERRORID : L_IE1P_Error;
	LRINPUTMAGNITUDE : LREAL;
	LRINPUTPHASE : LREAL;
	LROUTPUTMAGNITUDE : LREAL;
	LROUTPUTPHASE : LREAL;
	DWACTINDEX : DWORD;
	STRFORMATED : STRING(255);
END_VAR
VAR
	_ITFLOCKABLE : L_UBUP_ILockable;
	_MODEL : L_UBUP_BehaviourModel_ETrigA;
END_VAR
END_FUNCTION_BLOCK

METHOD CYCLICACTION
VAR_INPUT
	ITFTIMINGCONTROLLER : L_UBUP_ITimingController;
END_VAR
VAR_OUTPUT
	XCOMPLETE : BOOL;
	XABORT : BOOL;
	IERRORID : INT;
END_VAR
END_METHOD

METHOD FINALIZEACTION
VAR_INPUT
	XABORTPROPOSED : BOOL;
	IERRORIDPROPOSED : INT;
END_VAR
VAR_OUTPUT
	XCOMPLETE : BOOL;
	XABORT : BOOL;
	IERRORID : INT;
END_VAR
END_METHOD

METHOD RESETACTION
VAR_OUTPUT
	XCOMPLETE : BOOL;
END_VAR
END_METHOD

METHOD STARTACTION
VAR_OUTPUT
	XCOMPLETE : BOOL;
	IERRORID : INT;
END_VAR
END_METHOD
